(* IEC 61131-3 sources: daoli-st-library/DL_Motion (part 10) *)

(* ---- FB_DL_AxisTorqueRippleWatch.st ---- *)
(*
  Name        : FB_DL_AxisTorqueRippleWatch
  Category    : DL_Motion
  Version     : 1.0.0
  Purpose     : 轴转矩纹波监视：匀速段窗内峰峰值/均值占比与峰间隔规律性双判据，识别机械卡滞与联轴器异常；/ Axis torque ripple watch: peak-to-mean ripple ratio and peak-interval regularity in a steady-speed window to identify mechanical sticking and coupling anomalies
  溯源        : 借 plcopen-motion 的运动诊断组织，clean-room 实现
  Boundary    : ① 只在匀速段采样（|速度 - 速度命令| < 容差 且 速度 > 最低速），运动相位闸（容差/最低速域 > 0）；
                ② 波动幅度 = 窗内峰峰值 / 均值占比判据，均值近零时占比出口置 0 + bInvalid（除零前置）；
                ③ 周期性判据 = 峰间隔极差 < 阈（机械卡滞特征），需窗内 >= 3 个局部峰才判；
                ④ 非有限扭矩该拍不入窗（窗保持不滑动，防污染统计）；
                ⑤ 本件为诊断观测层，不干预轴指令输出（属主边界，零控制量引脚）；
                ⑥ 窗长 32 固定常量，窗内统计每趟全量重算防陈旧（R227）。
*)
TYPE E_DL_TrwState :
(
    eIdle  := 0,                             (* 未使能（窗清空） / Disabled, window cleared *)
    eRun   := 10,                            (* 纹波监视运行 / Watching *)
    eFault := 90                             (* 故障锁存相 / Fault latched *)
);
END_TYPE

TYPE E_DL_TrwCause :
(
    eNone      := 0,                         (* 无成因 / No cause *)
    eCfgIllegal:= 1,                        (* 组态非法：容差/最低速/阈值/周期越域 / Illegal config *)
    ePhaseBad  := 2                         (* 非法相位兜底 / Illegal phase fallback *)
);
END_TYPE

FUNCTION_BLOCK FB_DL_AxisTorqueRippleWatch
VAR_INPUT
    fTorque  : REAL := 0.0;                  (* 轴转矩反馈 [Nm] / Axis torque feedback *)
    fVel     : REAL := 0.0;                 (* 轴实际速度 [mm/s] / Actual velocity *)
    fVelCmd  : REAL := 0.0;                 (* 轴速度命令（匀速判据基准）[mm/s] / Velocity command *)
    fVelTol  : REAL := 5.0;                  (* 匀速判据容差，域 > 0 [mm/s] / Steady-speed tolerance *)
    fVelMin  : REAL := 10.0;                 (* 最低采样速度，域 > 0 [mm/s] / Minimum sampling speed *)
    fTqLimRip: REAL := 10.0;                 (* 纹波占比报警阈，域 > 0 [%] / Ripple ratio limit *)
    fGapSpreadMax: REAL := 0.05;             (* 峰间隔极差阈，域 > 0 [s] / Gap spread limit *)
    tSample  : TIME := T#10MS;               (* 采样周期，域 > T#0S [ms] / Sampling period *)
    bEnable  : BOOL := TRUE;                 (* 使能 [-] / Enable *)
    bReset   : BOOL := FALSE;                (* 复位命令，上升沿清窗与故障 [-] / Reset command *)
END_VAR
VAR_OUTPUT
    fRipplePct: REAL;                        (* 纹波占比出口 = 峰峰值 / |均值| × 100 [%] / Ripple ratio outlet *)
    bRippleHigh: BOOL;                       (* 纹波超阈判据出口 [-] / Ripple high verdict *)
    bPeriodic: BOOL;                         (* 周期性卡滞特征出口（>= 3 峰且间隔规律）[-] / Periodic sticking verdict *)
    bInvalid : BOOL;                         (* 本拍统计无效指示（均值近零/样本不足）[-] / Invalid indicator *)
    eState   : E_DL_TrwState;                (* 状态出口 / State outlet *)
    eCause   : E_DL_TrwCause;                (* 故障成因出口（R190 归因唯一） / Fault cause outlet *)
    bError   : BOOL;                         (* 故障锁存标志 [-] / Fault latch flag *)
END_VAR
VAR
    _eState : E_DL_TrwState := E_DL_TrwState.eIdle;  (* 内部相位（CASE 唯一写入目标） / Internal phase *)
    _eCause : E_DL_TrwCause := E_DL_TrwCause.eNone;  (* 成因锁存量 / Latched cause *)
    rtReset : R_TRIG;                        (* 复位沿实例，段 0 无条件调用 / Reset edge instance *)
    _bFault : BOOL;                          (* 故障锁存位 / Latched fault bit *)
    _bCfgBad: BOOL;                          (* 组态非法当拍量 / Illegal config this scan *)
    _bFin   : BOOL;                          (* 扭矩有限性当拍量（边界④） / Torque finiteness *)
    _bSteady: BOOL;                          (* 匀速段当拍判据（边界①） / Steady-speed verdict *)
    _aWin   : ARRAY[1..32] OF REAL;          (* 扭矩滑窗（线性平移式）[Nm] / Torque sliding window *)
    _nFill  : INT;                           (* 窗填充数 [点] / Window fill count *)
    _i      : INT;                           (* 窗扫描游标 [点] / Window scan cursor *)
    _fMean  : REAL;                          (* 窗均值中间量 [Nm] / Window mean *)
    _fPk    : REAL;                          (* 窗峰值中间量 [Nm] / Window peak *)
    _fTr    : REAL;                          (* 窗谷值中间量 [Nm] / Window trough *)
    _fSum   : REAL;                          (* 窗求和中间量 [Nm] / Window sum *)
    _nPkN   : INT;                           (* 本趟局部峰计数 [个] / Local peak count *)
    _nLastPk: INT;                           (* 上一峰样本序号（间隔派生）[点] / Last peak index *)
    _aGap   : ARRAY[1..4] OF REAL;           (* 最近峰间隔表（秒值）[s] / Recent peak gaps *)
    _nGapN  : INT;                           (* 已存间隔数 [个] / Stored gap count *)
    _fGapMax: REAL;                          (* 间隔极差上界中间量 [s] / Gap spread upper *)
    _fGapMin: REAL;                          (* 间隔极差下界中间量 [s] / Gap spread lower *)
    _fDtSec : REAL;                          (* 采样周期秒值，域 > eps [s] / Sampling period seconds *)
    _bPerI  : BOOL;                          (* 周期性判据内部量 / Periodic verdict internal *)
END_VAR
VAR CONSTANT
    DL_TRW_NMAX : INT   := 32;               (* 滑窗容量（固定常量，边界⑥）[点] / Window capacity *)
    DL_TRW_NMIN : INT   := 8;                (* 统计生效最少样本数（防小样本误判）[点] / Minimum samples *)
    DL_TRW_NPKMIN: INT  := 3;                (* 周期性判据最少峰数（边界③）[个] / Minimum peaks *)
    DL_TRW_EPS  : REAL  := 1.0E-6;           (* 判零容差 [-] / Epsilon *)
END_VAR

(* —— 段 0：当拍判据派生 + 实例无条件刷新（R228A） —— *)
_fDtSec := TIME_TO_LREAL(tSample) / 1000.0;              (* 采样周期秒化（除子常量 1000） / Sampling period seconds *)
_bCfgBad := (fVelTol <= DL_TRW_EPS) OR (fVelMin <= DL_TRW_EPS)           (* 匀速容差/最低速正域闸（边界①） / Tolerance and speed gates *)
            OR (fTqLimRip <= DL_TRW_EPS) OR (fGapSpreadMax <= DL_TRW_EPS)   (* 报警阈正域闸（边界②③） / Verdict limit gates *)
            OR NOT (tSample > T#0S);                     (* 采样周期正域闸 / Sampling gate *)
rtReset(CLK := bReset);                                  (* 复位沿每拍必调 / Reset edge every scan *)
_bFin := (fTorque = fTorque) AND ((fTorque - fTorque) = (fTorque - fTorque));   (* 扭矩 NaN 自反 + Inf 差判闸（边界④） / Torque NaN and Inf gate *)
_bSteady := (ABS(fVel - fVelCmd) < fVelTol) AND (fVel > fVelMin);        (* 匀速段判据：速度差容差内且高于最低速（边界①） / Steady-speed verdict *)

(* —— 段 1：单拍量预清零（R107；出口在段 4 每趟重算前预置确定值） —— *)
fRipplePct := 0.0;                                       (* 占比出口预清（无效拍默认 0） / Ripple preset zero *)
bRippleHigh := FALSE;                                    (* 超阈出口预清 / High preset *)
bPeriodic := FALSE;                                      (* 周期性出口预清 / Periodic preset *)
bInvalid := FALSE;                                       (* 无效指示预清 / Invalid preset *)
_bPerI := FALSE;                                         (* 周期性内部量预清（R227） / Periodic internal clear *)
_nPkN := 0;                                              (* 峰计数每趟重置 / Peak count reset *)
_nLastPk := 0;                                           (* 峰序号快照重置 / Peak index reset *)
_nGapN := 0;                                             (* 间隔表计数每趟重算 / Gap count reset *)
_fGapMax := 0.0;                                         (* 极差上界重置 / Spread upper reset *)
_fGapMin := 0.0;                                         (* 极差下界重置 / Spread lower reset *)

(* —— 段 2：复位沿处理（作用域：清故障 + 清窗 + 迁 eIdle，R283 逐项声明） —— *)
IF rtReset.Q THEN
    _bFault := FALSE;                                    (* 清故障锁存 / Clear fault *)
    _eCause := E_DL_TrwCause.eNone;                      (* 清成因 / Clear cause *)
    FOR _i := 1 TO DL_TRW_NMAX DO
        _aWin[_i] := 0.0;                                (* 清滑窗 / Clear window *)
    END_FOR
    FOR _i := 1 TO 4 DO
        _aGap[_i] := 0.0;                                (* 清间隔表 / Clear gap table *)
    END_FOR
    _nFill := 0;                                         (* 清窗填充数 / Clear fill *)
    fRipplePct := 0.0;                                   (* 清占比出口 / Clear ripple outlet *)
    _eState := E_DL_TrwState.eIdle;                      (* 迁未使能相 / Back to idle *)
END_IF

(* —— 段 3：组态故障锁存（锁存至复位沿，R189） —— *)
IF _bCfgBad AND NOT _bFault THEN
    _bFault := TRUE;                                     (* 锁存故障位 / Latch fault *)
    _eCause := E_DL_TrwCause.eCfgIllegal;                (* 成因：组态非法 / Cause illegal config *)
    _eState := E_DL_TrwState.eFault;                     (* 同步迁故障相 / Migrate to fault *)
END_IF

(* —— 段 4：CASE 主状态机（ELSE 兜底迁 eFault，红线 6） —— *)
CASE _eState OF
    E_DL_TrwState.eIdle:                                 (* 未使能：窗清空出口确定值 / Idle *)
        FOR _i := 1 TO DL_TRW_NMAX DO
            _aWin[_i] := 0.0;                            (* 失能清滑窗 / Disabled clear window *)
        END_FOR
        _nFill := 0;                                     (* 失能清填充数 / Disabled clear fill *)
        IF bEnable AND NOT _bFault THEN
            _eState := E_DL_TrwState.eRun;               (* 进入监视相 / Enter watching *)
        END_IF
    E_DL_TrwState.eRun:                                  (* 监视相：匀速闸采样 + 全窗重算 / Watching *)
        IF NOT bEnable THEN
            _eState := E_DL_TrwState.eIdle;              (* 失能回未使能 / Back to idle *)
        ELSE
            IF _bSteady AND _bFin AND (_fDtSec > DL_TRW_EPS) THEN   (* 匀速闸 + 有限闸 + 周期闸（边界①④） / Sampling gates *)
                IF _nFill < DL_TRW_NMAX THEN
                    _nFill := _nFill + 1;                (* 填充数递进（写入点域内） / Fill advance *)
                    _aWin[_nFill] := fTorque;            (* 样本入窗 / Sample into window *)
                ELSE
                    FOR _i := 1 TO DL_TRW_NMAX - 1 DO
                        _aWin[_i] := _aWin[_i + 1];      (* 满窗线性平移（有界循环） / Shift window *)
                    END_FOR
                    _aWin[DL_TRW_NMAX] := fTorque;       (* 新样本入窗尾 / Sample into tail *)
                END_IF
            END_IF                                       (* 不满足闸：本拍不入窗（窗保持，边界①④） *)
            IF _nFill >= DL_TRW_NMIN THEN                (* 统计生效下限（防小样本误判） / Statistics gate *)
                _fSum := 0.0; _fPk := _aWin[1]; _fTr := _aWin[1];   (* 均值/峰谷初值（R227） / Init mean peak trough *)
                FOR _i := 1 TO _nFill DO
                    _fSum := _fSum + _aWin[_i];          (* 窗求和 / Window sum *)
                    IF _aWin[_i] > _fPk THEN
                        _fPk := _aWin[_i];               (* 窗峰值刷新 / Peak update *)
                    END_IF
                    IF _aWin[_i] < _fTr THEN
                        _fTr := _aWin[_i];               (* 窗谷值刷新 / Trough update *)
                    END_IF
                END_FOR
                _fMean := _fSum / INT_TO_REAL(_nFill);   (* 窗均值（除子 = 填充数 >= 8） / Window mean *)
                IF ABS(_fMean) > DL_TRW_EPS THEN
                    fRipplePct := (_fPk - _fTr) / ABS(_fMean) * 100.0;   (* 纹波占比（除子已过闸，边界②） / Ripple ratio *)
                    bRippleHigh := fRipplePct > fTqLimRip;   (* 占比超阈判据（直比阈值） / Ripple high verdict *)
                ELSE
                    fRipplePct := 0.0;                   (* 均值近零：占比出口 0（除零前置，边界②） / Zero ratio *)
                    bInvalid := TRUE;                    (* 无效指示 / Invalid indicator *)
                END_IF
                FOR _i := 2 TO _nFill - 1 DO             (* 局部峰检测（内点扫描，边界③） / Local peak scan *)
                    IF (_aWin[_i] > _aWin[_i - 1]) AND (_aWin[_i] > _aWin[_i + 1]) AND (_aWin[_i] > _fMean) THEN
                        _nPkN := _nPkN + 1;              (* 局部峰计数 / Peak count *)
                        IF _nLastPk >= 1 THEN
                            _nGapN := _nGapN + 1;        (* 间隔数净额 +1 / Gap count *)
                            IF _nGapN > 4 THEN
                                _aGap[1] := _aGap[2]; _aGap[2] := _aGap[3]; _aGap[3] := _aGap[4];   (* 间隔表平移 / Shift gaps *)
                                _nGapN := 4;             (* 间隔表封顶 / Gap cap *)
                            END_IF
                            _aGap[_nGapN] := INT_TO_REAL(_i - _nLastPk) * _fDtSec;   (* 间隔秒值入表 / Gap into table *)
                        END_IF
                        _nLastPk := _i;                  (* 峰序号快照 / Peak index snapshot *)
                    END_IF
                END_FOR
                IF _nGapN >= 2 THEN                      (* >= 3 峰（2 个间隔）才判（边界③） / Peak count gate *)
                    _fGapMax := _aGap[1]; _fGapMin := _aGap[1];   (* 极差初值 / Spread init *)
                    FOR _i := 2 TO _nGapN DO
                        IF _aGap[_i] > _fGapMax THEN
                            _fGapMax := _aGap[_i];       (* 间隔上界刷新 / Gap upper *)
                        END_IF
                        IF _aGap[_i] < _fGapMin THEN
                            _fGapMin := _aGap[_i];       (* 间隔下界刷新 / Gap lower *)
                        END_IF
                    END_FOR
                    _bPerI := (_fGapMax - _fGapMin) < fGapSpreadMax;   (* 间隔规律性判据（边界③） / Regularity verdict *)
                END_IF
                bPeriodic := _bPerI;                     (* 周期性出口 / Periodic outlet *)
            ELSE
                bInvalid := TRUE;                        (* 样本不足：统计无效（确定值） / Not enough samples *)
            END_IF
        END_IF
    E_DL_TrwState.eFault:                                (* 故障相：冻结保持，仅复位沿出 / Fault *)
        ;                                                (* 锁存回放（R28） / Replay from latch *)
    ELSE                                                 (* 非法相位兜底迁安全态 / Illegal phase fallback *)
        _eState := E_DL_TrwState.eFault; _bFault := TRUE;    (* 迁故障相 + 同步锁存 / To fault and latch *)
        _eCause := E_DL_TrwCause.ePhaseBad;              (* 成因：非法相位 / Cause illegal phase *)
END_CASE

(* —— 段 5：出口映射（bError/eState 同源，R191） —— *)
bError := _bFault;                                       (* 故障标志镜像 / Fault flag mirror *)
eState := _eState;                                       (* 状态出口 / State outlet *)
eCause := _eCause;                                       (* 成因出口 / Cause outlet *)
END_FUNCTION_BLOCK

(* ---- FB_DL_AxisTorqueWatch.st ---- *)
(*
  组件名 Component   : FB_DL_AxisTorqueWatch
  子库 Sublibrary    : DL_Motion
  版本 Version       : 1.0.0
  兼容性 Platform    : CODESYS 3.5 / TwinCAT 3 / 汇川 InoProShop / Machine Expert（仅 Standard.library）
  功能 Function      : 轴转矩趋势监视（与 FB_DL_TorqueLimitControl 分工：控 vs 监）：
                       1) 带域判据：转矩超上带限持续 tConfirmWin → 预警（bWarn）；
                       2) 趋势斜率判据：周期窗（tSlopeWin 自复触）两端采样，斜率
                       fSlopeNmS = (本端 - 上端) / 窗长，斜率超限 → 预警；
                       3) 堵转分级：转矩超上带限 且 轴速近零 持续 tStallTo → bStall；
                       4) 三判据各带独立确认窗，互不共用计时实例（R190 归因唯一）。
  边界 Boundary      : ① 监视件只出分级诊断位，不接管转矩控制输出；
                       ② 周期窗计时用 IN := bEnable AND NOT tonSlopeWin.Q 自复触
                       （R188 错峰周期窗范式，禁外部沿清零）；
                       ③ 斜率除法前置域闸：tSlopeWin <= T#0S 判组态非法；
                       ④ 非有限值（NaN 自反 + 无穷差值自减）判输入非法锁存；
                       ⑤ 故障锁存解除唯一路径 = bReset 上升沿（输入引脚，恒可达）；
                       ⑥ 无全局变量引用、无外部变量声明、无物理地址寻址。
  依赖 Depends       : Standard.library（R_TRIG / TON）
  溯源 Origin        : 道莅自研 clean-room（参考 t2-4-s7-motion 监视分类与参数域，
                       零代码行复制）
  码位 Code          : 16#04_0_A9
  码表 Error codes（Motion 格 04_0_A9，单轨：故障 0x02A9 / 信息 0x01A9 / 0x03A9）:
    16#0004_02A9 故障级：组态非法或输入非有限，锁存至 bReset 上升沿
    16#0004_01A9 信息级：预警进入沿（bWarn 由 FALSE 转 TRUE 拍）
    16#0004_05A9 信息级：堵转检出沿（bStall 由 FALSE 转 TRUE 拍；子道 05 为 03 道撞车顺延勘误）
  修订历史 Revision  :
    2026-11-19  v1.0.0  R44 首版（批次 2 · 序号 6）
*)

TYPE E_DL_AtwState :
(
    eIdle  := 0,    // 空闲：未使能 / Idle, not enabled
    eRun   := 10,   // 监视运行：三判据并行 / Running, three criteria active
    eFault := 90    // 故障：组态/输入锁存 / Fault, latched
);
END_TYPE

FUNCTION_BLOCK FB_DL_AxisTorqueWatch
VAR_INPUT
    bEnable    : BOOL;                     // 使能（电平）[-] / Enable
    bReset     : BOOL;                     // 上升沿清故障锁存 [-] / Reset edge
    fTorqueNm  : REAL;                     // 实测转矩 [牛·米] / Measured torque
    fVelMmS    : REAL;                     // 轴实际速度 [mm/s] / Axis velocity
    fBandHiNm  : REAL := 10.0;             // 转矩上带限 [牛·米] / Torque band ceiling
    fBandLoNm  : REAL := 1.0;              // 转矩下带限 [牛·米] / Torque band floor
    fSlopeLimNmS: REAL := 5.0;             // 趋势斜率限值 [牛·米/秒] / Trend slope limit
    fVelNearZeroMmS: REAL := 0.5;          // 堵转判近零速度阈 [mm/s] / Near-zero velocity threshold
    tConfirmWin: TIME := T#2S;             // 带域预警确认窗 [毫秒] / Band confirm window
    tSlopeWin  : TIME := T#1S;             // 趋势斜率测量窗 [毫秒] / Slope measurement window
    tStallTo   : TIME := T#3S;             // 堵转确认窗 [毫秒] / Stall confirm window
END_VAR
VAR_OUTPUT
    bInBand    : BOOL;                     // 转矩在带内电平 [-] / Torque in-band level
    bWarn      : BOOL;                     // 预警电平（带域或斜率越限确认后）[-] / Warning level
    bStall     : BOOL;                     // 堵转电平 [-] / Stall level
    fSlopeNmS  : REAL;                     // 实测趋势斜率 [牛·米/秒] / Measured slope
    eState     : E_DL_AtwState;            // 状态出口，段尾单点映射 / State outlet
    bError     : BOOL;                     // 故障锁存标志 [-] / Fault latch flag
    uErrId     : UDINT;                    // 事件码，0 = 无事件 / Event code
END_VAR
VAR
    rtReset    : R_TRIG;                   // 复位沿实例，段 0 无条件刷新 / Reset edge
    rtWarn     : R_TRIG;                   // 预警进入沿实例，段 0 无条件刷新 / Warn entry edge
    rtStall    : R_TRIG;                   // 堵转进入沿实例，段 0 无条件刷新 / Stall entry edge
    tonBandWin : TON;                      // 带域确认窗（专用确认窗命名） / Band confirm timer
    tonStallTo : TON;                      // 堵转确认窗（专用超时件命名（R228A 豁免）） / Stall timer
    tonSlopeWin: TON;                      // 斜率周期窗（自复触，R188） / Slope window timer
    _eState    : E_DL_AtwState := E_DL_AtwState.eIdle;   // 内部相位（CASE 唯一写入目标）/ Internal phase
    _bBandHi   : BOOL;                     // 带域越限当拍量 [-] / Band breach flag
    _bStallCond: BOOL;                     // 堵转条件当拍量 [-] / Stall condition flag
    _fTorqueSnap: REAL;                    // 窗始转矩快照 [牛·米] / Window-start torque snapshot
    _bSnapPend : BOOL;                     // 快照待取标志 [-] / Snapshot pending flag
    _bFault    : BOOL;                     // 故障锁存位（锁存量） / Latched fault bit
    _uFault    : UDINT;                    // 故障码锁存（锁存量） / Latched fault code
    _bCfgBad   : BOOL;                     // 组态非法当拍量 [-] / Config illegal flag
    _bNonFin   : BOOL;                     // 输入非有限当拍量 [-] / Non-finite input flag
END_VAR
VAR CONSTANT
    DL_SLOPE_EPS: REAL := 1.0E-9;          // 斜率判零容差 [牛·米/秒] / Slope tolerance
    DL_WIN_EPS  : REAL := 1.0E-3;          // 窗长秒值下限 [秒] / Window seconds floor
    DL_ABS_MAX  : REAL := 1.0E30;          // 有限值判定上界 [工程单位] / Finite bound
    DL_ZERO     : REAL := 0.0;             // 零常量 [工程单位] / Zero constant
    DL_MS_PER_S : REAL := 1000.0;          // 毫秒 → 秒换算系数 [毫秒/秒] / Milliseconds per second
END_VAR

(* —— 段 0｜沿与定时器每拍无条件刷新（禁置于 IF/CASE 内） —— *)
_bBandHi    := (fTorqueNm > fBandHiNm) OR (fTorqueNm < fBandLoNm);   // 带域越限当拍判据
_bStallCond := (fTorqueNm > fBandHiNm) AND (ABS(fVelMmS) < fVelNearZeroMmS);
rtReset    (CLK := bReset);
rtWarn     (CLK := bWarn);
rtStall    (CLK := bStall);
tonBandWin (IN := (_eState = E_DL_AtwState.eRun) AND _bBandHi AND (NOT _bFault), PT := tConfirmWin);
tonStallTo (IN := (_eState = E_DL_AtwState.eRun) AND _bStallCond AND (NOT _bFault), PT := tStallTo);
tonSlopeWin(IN := (_eState = E_DL_AtwState.eRun) AND (NOT _bFault) AND (NOT tonSlopeWin.Q),
            PT := tSlopeWin);            // 自复触周期窗：Q 拍断开一拍，下拍重启（R188）

(* —— 段 1｜瞬时量预清零（锁存量 _bFault/_uFault/bWarn/bStall/_fTorqueSnap 不入清单） —— *)
uErrId   := 16#0000_0000;
_bCfgBad := FALSE;
_bNonFin := FALSE;

(* —— 段 2｜复位沿：故障一次性清干净，相位回空闲，诊断位复归 —— *)
IF rtReset.Q THEN
    _bFault  := FALSE;
    _uFault  := 16#0000_0000;
    bWarn    := FALSE;
    bStall   := FALSE;
    fSlopeNmS:= DL_ZERO;
    _eState  := E_DL_AtwState.eIdle;
END_IF

(* —— 段 3｜组态闸与非有限判据 —— *)
IF (fBandHiNm <= fBandLoNm) OR (tConfirmWin = T#0S) OR (tSlopeWin = T#0S)
   OR (tStallTo = T#0S) OR (fVelNearZeroMmS <= DL_ZERO) THEN
    _bCfgBad := TRUE;
END_IF
IF (fTorqueNm <> fTorqueNm) OR ((fTorqueNm - fTorqueNm) <> DL_ZERO)
   OR (fVelMmS <> fVelMmS) OR ((fVelMmS - fVelMmS) <> DL_ZERO) THEN
    _bNonFin := TRUE;
END_IF

(* —— 段 4｜主状态机：三态全覆盖 + ELSE 兜底 —— *)
CASE _eState OF

E_DL_AtwState.eIdle:
    bInBand := FALSE;
    IF bEnable AND (NOT _bCfgBad) AND (NOT _bNonFin) THEN
        _fTorqueSnap := fTorqueNm;       // 窗始快照初始化
        _bSnapPend   := FALSE;
        _eState := E_DL_AtwState.eRun;
    ELSIF bEnable AND (_bCfgBad OR _bNonFin) THEN
        _bFault := TRUE;
        _uFault := 16#0004_02A9;
        bError  := TRUE;
        _eState := E_DL_AtwState.eFault;
    END_IF

E_DL_AtwState.eRun:
    IF NOT bEnable THEN
        bInBand := FALSE;
        bWarn   := FALSE;
        bStall  := FALSE;
        _eState := E_DL_AtwState.eIdle;  // 使能撤销回空闲
    ELSE
        bInBand := NOT _bBandHi;
        (* 斜率测量：Q 拍收口，快照按窗复归（除数 = 窗长秒值，组态闸已保证 > 0） *)
        IF tonSlopeWin.Q THEN
            IF NOT _bSnapPend THEN
                fSlopeNmS := (fTorqueNm - _fTorqueSnap)
                             / MAX(TIME_TO_REAL(tSlopeWin) / DL_MS_PER_S, DL_WIN_EPS);
                IF ABS(fSlopeNmS) < DL_SLOPE_EPS THEN
                    fSlopeNmS := DL_ZERO;    // 斜率近零归零
                END_IF
                _bSnapPend := TRUE;
            END_IF
            _fTorqueSnap := fTorqueNm;
            _bSnapPend   := FALSE;
        END_IF
        (* 分级判据：带域或斜率任一确认 → 预警；带域 + 近零速度确认 → 堵转 *)
        IF _bNonFin THEN
            _bFault := TRUE;             // 输入非有限：运行中锁存
            _uFault := 16#0004_02A9;
            bError  := TRUE;
            bWarn   := FALSE;
            bStall  := FALSE;
            _eState := E_DL_AtwState.eFault;
        ELSE
            bWarn := (NOT _bFault) AND (tonBandWin.Q OR (ABS(fSlopeNmS) > fSlopeLimNmS));
            bStall := (NOT _bFault) AND tonStallTo.Q;
            IF rtWarn.Q THEN
                uErrId := 16#0004_01A9;  // 信息级：预警进入沿
            END_IF
            IF rtStall.Q THEN
                uErrId := 16#0004_05A9;  // 信息级：堵转检出沿（子道 05 勘误顺延）
            END_IF
        END_IF
    END_IF

E_DL_AtwState.eFault:
    bError := TRUE;                      // 故障相驻留：诊断位冻结，只认复位沿（段 2 迁出）
    ;                                    // （冻结语义：bWarn/bStall 保持复位沿前值由段 2 归零）

ELSE
    _bFault := TRUE;                     // 兜底：非法相位锁存
    _uFault := 16#0004_02A9;
    bError  := TRUE;
    _eState := E_DL_AtwState.eFault;
END_CASE

(* —— 段 5｜状态出口单点映射 —— *)
eState := _eState;
END_FUNCTION_BLOCK

(* ---- FB_DL_AxisVelocityMove.st ---- *)
(*==============================================================================
 * 组件名称 (Component)  : FB_DL_AxisVelocityMove
 * 所属子库 (Sublibrary) : DL_Motion
 * 当前版本 (Version)    : 1.0.0
 * 组件分类 (Category)   : 功能块（FUNCTION_BLOCK）· 单轴速度模式与动态变速封装 · 工艺上层件
 * 兼容性   (Platform)   : CODESYS 3.5 / TwinCAT 3 / 汇川 InoProShop / Schneider
 *                         Machine Expert；仅依赖 Standard.library（R_TRIG /
 *                         F_TRIG / MIN / MAX / ABS），零厂商方言
 * 接口依赖 (Depends)    : I_DL_MotionAxis / E_DL_AxisState（既有契约，Round 05）
 * 功能描述 (Function)   : 单轴速度模式（MC_MoveVelocity 语义）与动态变速控制
 *                         封装。经轴接口引用驱动轴体：指令电平生效，TRUE=运行
 *                         / FALSE=受控停止；运行中变更 fVelocity 即为改速请求
 *                         （轴接口连续运动改速语义，改速而非重启），bDynamicRetarget
 *                         使能时自动重发；速度上限独立钳位，越限置信息级。
 * 设计要点 (Key notes)  : ① 指令上升沿门禁：轴待机态受理运行、连续运动态受理
 *                           改速；其余态请求不被受理 → 信息级 0004_0107；
 *                         ② 动态改速：连续运动中 |fVelocity − 上次已发值| 超
 *                           容差即重发 MoveVelocity（改速语义），指令被拒 →
 *                           0004_0230 故障级锁存；
 *                         ③ 下降沿 → 轴受控停止（MC_Stop 语义）；
 *                         ④ 参数门禁（fAcc 非正值/非有限值）→ 信息级 0004_0106
 *                           （与 FB_DL_AxisHomingSeq/FB_DL_AxisRelativeMove
 *                           同码同义：参数门禁拒绝，共用留档）；
 *                         ⑤ 本块为事件型 + 轮询状态组件，免首扫（R23）。
 * 开源溯源 (Origin)     : 原创实现（参考 PLCopen Part 1-6 MC_MoveVelocity 公开
 *                         语义与西门子 Motion Control 对象语义，clean-room）。
 *                         仅提取公开指令动词、参数域与改速语义；实现与命名
 *                         100% 自有，未参考任何厂商源码行。
 * 验收向量 (Acceptance) :
 *   V1 启动-停止链：bCmdStart 上升沿→轴进连续运动；下降沿→受控停止；
 *   V2 运行中改速：fVelocity 50→-30（含反向）→ 自动重发改速，轴不重启；
 *   V3 改速被拒：轴受控停止中发改速请求 → 信息级 0004_0107，轴不受扰；
 *   V4 速度钳位：|fVelocity|=5000 > fVelMax=1000 → 钳位至 1000 + 信息级；
 *   V5 轴故障中断：运行中轴故障反馈 → 0004_0230 锁存，bBusy 退出。
 * 故障码表 (Error codes):
 *   16#0004_0106【信息级】参数门禁拒绝（三块同码同义，共用留档）；
 *   16#0004_0107【信息级】改速请求不被受理/速度钳位提示（规格外补充子义，
 *   R11 留档）；16#0004_0230【故障级】指令被拒/轴故障中断（锁存）；
 *   16#0004_0201【故障级】非法状态兜底（沿用族码，与 FB_DL_SingleAxis 同码
 *   同义，复用留档）。
 * 修订历史 (Revision)   :
 *   2026-11-15  v1.0.0  首版入库（Round 06 · DL_Motion 回零/运动族）
 *============================================================================*)

(*-----------------------------------------------------------------------------
 * 调用示例 (Instance guide)：
 *   fbVel.iAxis := fbAxis;                        // 接口依赖注入
 *   fbVel(bCmdStart := bRunSwitch, fVelocity := fSetVel, // 周期调用
 *         fAcc := 2000.0, bDynamicRetarget := TRUE, fVelMax := 1000.0);
 *   电平语义：bRunSwitch 断开即受控减速停车，无需上层编排停止时序；
 *   改速只需改 fVelocity 输入值，块自动差值比较后重发改速指令。
 *----------------------------------------------------------------------------*)

(*-----------------------------------------------------------------------------
 * 常见误用与现场提示 (Field notes)：
 *   1 bCmdStart 电平语义：FALSE 即停车并退出速度模式，不要用脉冲；
 *     需要脉冲语义的工位在上层自锁存。
 *   2 改速容差为固定值（0.001 mm/s），HMI 微调速度时每次变化都会重发；
 *     高频改速场景请在上层做死区滤波，避免指令流量放大。
 *   3 轴限位停车后 bCmdStart 仍为 TRUE 时本块会自动重新发起（电平需求
 *     语义）；不希望自动重启的工位在限位联动层断开 bCmdStart。
 *----------------------------------------------------------------------------*)

(*-----------------------------------------------------------------------------
 * 枚举: E_DL_VelStep（归属 DL_Motion，与 FB_DL_AxisVelocityMove 同文件）
 * 含义: 速度模式内部步进枚举（本块私有配套，外部仅作诊断参考）。
 *----------------------------------------------------------------------------*)
{attribute 'strict'}
{attribute 'qualified_only'}
TYPE E_DL_VelStep :
(
    eIdle    := 0,    // 空闲：等待启动沿 / Idle: waiting for start edge
    eRunning := 10    // 运行：轮询轴状态并处理动态改速 / Running: polling axis and retargeting
) UINT;
END_TYPE

FUNCTION_BLOCK FB_DL_AxisVelocityMove
VAR_INPUT
    bCmdStart        : BOOL := FALSE;   // 速度运行指令（Velocity start command），电平生效：TRUE=运行 / FALSE=受控停止
    fVelocity        : REAL := 0.0;     // 目标速度（Target velocity）[mm/s]，带符号，负值=负向；运行中变更即为改速请求
    fAcc             : REAL := 1000.0;  // 加减速度（Acceleration）[mm/s²]，正值，默认 1000.0
    bDynamicRetarget : BOOL := FALSE;   // 动态改速使能（Dynamic retarget），TRUE=连续运动中速度变化自动改速
    fVelMax          : REAL := 1000.0;  // 速度上限（Velocity limit）[mm/s]，|fVelocity| 超限钳位并置信息级
END_VAR
VAR_IN_OUT
    iAxis            : I_DL_MotionAxis; // 轴接口引用（Axis reference），由上层注入实现块实例
END_VAR
VAR_OUTPUT
    bBusy            : BOOL := FALSE;   // 速度模式激活（Velocity mode active）
    bActive          : BOOL := FALSE;   // 轴处于连续运动态（Axis in continuous motion），轮询派生
    uErrorId         : UDINT := 0;      // 末次事件码（Last error code），段位 16#0004_xxxx
END_VAR
VAR
    eStep            : E_DL_VelStep := E_DL_VelStep.eIdle; // 内部步进状态（Internal step state）
    bFaultLatch      : BOOL := FALSE;   // 故障锁存标志（Fault latch），0004_0230 锁存载体
    bParamOk         : BOOL := FALSE;   // 参数门禁通过标志（Parameter gate pass flag），逐拍重算
    fVelEff          : REAL := 0.0;     // 本拍钳位后的目标速度（Clamped target velocity）[mm/s]
    fVelSent         : REAL := 0.0;     // 上次已发轴指令速度（Last issued velocity）[mm/s]，改速差值比较基准
    fVelLim          : REAL := 1000.0;  // 生效速度上限（Effective velocity limit）[mm/s]，非有限值兜底
    fAccEff          : REAL := 1000.0;  // 生效加减速度（Effective acceleration）[mm/s²]，防除零兜底
    rtrigStart       : R_TRIG;          // 启动指令上升沿（Rising edge of start command）
    ftrigStart       : F_TRIG;          // 启动指令下降沿（Falling edge of start command）
END_VAR
VAR CONSTANT
    DL_VEL_INF_MAX   : REAL := 1.0E30;  // 有限值判定幅值上限（Finite-value magnitude bound）[mm/s 或 mm/s²]
    DL_VEL_EPS       : REAL := 1.0E-6;  // 浮点判零容差（Float zero tolerance）
    DL_VEL_TGT_TOL   : REAL := 1.0E-3;  // 改速差值容差（Retarget delta tolerance）[mm/s]，超过才重发改速
    DL_VEL_PAR_FLOOR : REAL := 1.0E-3;  // 加速度参数下限（Acceleration floor）[mm/s²]
END_VAR

// 段 1｜沿检测无条件周期刷新（R7 红线，严禁置于分支内）
rtrigStart(CLK := bCmdStart);
ftrigStart(CLK := bCmdStart);

// 段 2｜接口引用有效性防御：未注入轴引用则清输出退出（不产生误动作）
IF iAxis = 0 THEN
    bBusy := FALSE;
    bActive := FALSE;
    RETURN;
END_IF

// 段 3｜参数门禁逐拍重算（公约 0.8）：非法仅封锁启动（信息级 0004_0106），运行中不中断
bParamOk := (fAcc = fAcc) AND (fAcc <= DL_VEL_INF_MAX) AND (fAcc > DL_VEL_PAR_FLOOR);
IF (fVelMax = fVelMax) AND (fVelMax > DL_VEL_PAR_FLOOR) AND (fVelMax <= DL_VEL_INF_MAX) THEN
    fVelLim := fVelMax;                          // 合法速度上限直通 [mm/s]
ELSE
    fVelLim := 1000.0;                           // 非法上限兜底 [mm/s]
    uErrorId := 16#0004_0106;                    // 信息级：参数兜底修复提示
END_IF
fAccEff := MAX(fAcc, DL_VEL_PAR_FLOOR);          // 生效加速度下限兜底 [mm/s²]，防除零

// 段 4｜事件码管理（R15）：瞬时码逐拍重算，锁存码仅在新启动沿解除
IF NOT bFaultLatch THEN
    uErrorId := 0;
END_IF

// 段 5｜下降沿受控停车（电平语义：FALSE=停止；全局处理，任何态均生效）
IF ftrigStart.Q THEN
    iAxis.Stop();                                // 受控减速停车（MC_Stop 语义）
    bBusy := FALSE;
    IF eStep = E_DL_VelStep.eRunning THEN
        eStep := E_DL_VelStep.eIdle;             // 退出速度模式，等待下次启动沿
    END_IF
END_IF

// 段 6｜运行中轴故障中断（优先于状态机，锁存 R15）
IF (eStep = E_DL_VelStep.eRunning) AND iAxis.bError THEN
    bFaultLatch := TRUE;                         // 故障级锁存，仅新启动沿解除
    uErrorId := 16#0004_0230;
    bBusy := FALSE;
    eStep := E_DL_VelStep.eIdle;
END_IF

// 段 7｜速度模式状态机（ENUM + CASE + ELSE 兜底）
CASE eStep OF

    E_DL_VelStep.eIdle:                          // 空闲态：等待启动沿与门禁
        bBusy := FALSE;
        IF rtrigStart.Q THEN
            bFaultLatch := FALSE;                // 新启动沿：锁存码解除路径（R15）
            IF NOT bParamOk THEN
                uErrorId := 16#0004_0106;        // 参数门禁拒绝（信息级）
            ELSIF (iAxis.eState <> E_DL_AxisState.eStandstill)
              AND (iAxis.eState <> E_DL_AxisState.eContinuousMotion) THEN
                uErrorId := 16#0004_0107;        // 非受理态（停止中/故障态）：请求不被受理（信息级）
            ELSE
                fVelEff := fVelocity;            // 目标速度初值 [mm/s]
                IF fVelEff > fVelLim THEN
                    fVelEff := fVelLim;          // 正向超限钳位 [mm/s]
                    uErrorId := 16#0004_0107;    // 信息级：速度钳位提示
                ELSIF fVelEff < -fVelLim THEN
                    fVelEff := -fVelLim;         // 负向超限钳位 [mm/s]
                    uErrorId := 16#0004_0107;    // 信息级：速度钳位提示
                END_IF
                IF (fVelEff <> fVelEff) OR (ABS(fVelEff) > DL_VEL_INF_MAX) THEN
                    fVelEff := 0.0;              // 非有限速度防御归零（0=原地保持，安全侧）
                    uErrorId := 16#0004_0106;    // 信息级：参数门禁拒绝
                END_IF
                IF iAxis.MoveVelocity(fVelEff, fAccEff) THEN
                    fVelSent := fVelEff;         // 记录已发速度，作为改速差值基准 [mm/s]
                    eStep := E_DL_VelStep.eRunning;
                    bBusy := TRUE;
                ELSE
                    bFaultLatch := TRUE;         // 指令被轴拒绝：故障级锁存
                    uErrorId := 16#0004_0230;
                END_IF
            END_IF
        END_IF

    E_DL_VelStep.eRunning:                       // 运行态：电平需求语义 + 动态改速
        bBusy := TRUE;
        IF bCmdStart THEN
            fVelEff := fVelocity;                // 目标速度初值 [mm/s]
            IF fVelEff > fVelLim THEN
                fVelEff := fVelLim;              // 正向超限钳位 [mm/s]
                uErrorId := 16#0004_0107;        // 信息级：速度钳位提示
            ELSIF fVelEff < -fVelLim THEN
                fVelEff := -fVelLim;             // 负向超限钳位 [mm/s]
                uErrorId := 16#0004_0107;        // 信息级：速度钳位提示
            END_IF
            IF (fVelEff <> fVelEff) OR (ABS(fVelEff) > DL_VEL_INF_MAX) THEN
                fVelEff := 0.0;                  // 非有限速度防御归零（安全侧：请求停车速度）
                uErrorId := 16#0004_0106;        // 信息级：参数门禁拒绝
            END_IF
            IF iAxis.eState = E_DL_AxisState.eStandstill THEN
                // 轴已回待机（如限位自动停车）而需求电平仍为真：按电平需求重新发起
                IF iAxis.MoveVelocity(fVelEff, fAccEff) THEN
                    fVelSent := fVelEff;
                ELSE
                    bFaultLatch := TRUE;         // 重发被拒：故障级锁存
                    uErrorId := 16#0004_0230;
                    bBusy := FALSE;
                    eStep := E_DL_VelStep.eIdle;
                END_IF
            ELSIF bDynamicRetarget AND (ABS(fVelEff - fVelSent) > DL_VEL_TGT_TOL) THEN
                // 动态改速：连续运动中差值超容差 → 重发改速（改速而非重启，接口契约语义）
                IF iAxis.eState = E_DL_AxisState.eContinuousMotion THEN
                    IF iAxis.MoveVelocity(fVelEff, fAccEff) THEN
                        fVelSent := fVelEff;     // 更新已发速度基准 [mm/s]
                    ELSE
                        bFaultLatch := TRUE;     // 改速指令被拒：故障级锁存
                        uErrorId := 16#0004_0230;
                        bBusy := FALSE;
                        eStep := E_DL_VelStep.eIdle;
                    END_IF
                ELSE
                    uErrorId := 16#0004_0107;    // 改速请求在非受理态被拒（信息级，瞬态）
                END_IF
            END_IF
        END_IF

    ELSE
        // 非法状态兜底（故障级，沿用族码 0004_0201，复用留档）
        uErrorId := 16#0004_0201;
        bFaultLatch := TRUE;
        bBusy := FALSE;
        eStep := E_DL_VelStep.eIdle;

END_CASE

// 段 8｜状态出口派生（R21：bActive 为轴状态轮询派生式，逐拍重算）
bActive := (iAxis.eState = E_DL_AxisState.eContinuousMotion);
END_FUNCTION_BLOCK

(* ---- FB_DL_BacklashCompensator.st ---- *)
(*
    FB_DL_BacklashCompensator —— 换向背隙补偿
    ------------------------------------------------------------------
    分类      : DL_Motion / Compensation
    前缀      : FB_DL_
    版本      : 1.0.1
    溯源      : T1-6 轴级补偿语义（只借「换向补偿属运动层给定量修正」的分类事实）；
                T2-2 LBP 泵 / 辊「背隙两阶段逼近」组织方式为次源（该组织已被
                RollerGapAdjust 使用）；增量式补偿、EWMA 学习、容差闸与码位 100% 自有；
                clean-room 重写，未复制任何闭源厂商源码，参考实现仅限 MIT/Apache 许可
    平台      : 纯 IEC 61131-3，CODESYS V3.5+ / TwinCAT 3 / InoProShop 通用
    作者      : 道莅代码库 · PLC编程专家（R18）
    ------------------------------------------------------------------
    功能说明  : 指令方向翻转瞬间在给定量上叠加一个方向性补偿量，抵消齿轮 / 丝杠反向
                间隙；并在到位后按实测偏差用 EWMA 自学习背隙估计（现场背隙随磨损变化）；
                与 FB_DL_RollerGapAdjust 的分界是后者为工艺辊缝调整顺控，本件是轴级
                给定量修正，两者不重叠；
                三道闸：负背隙取绝对值（参数习惯差异，不是故障）→ 超上限判故障
                （10 mm 以上补偿会把轴推到撞块）→ 位置非有限即旁路并清方向记忆；
                方向判定带死区，浮点判等全部带容差，杜绝边界来回翻转导致的补偿抖动；
                首拍没有历史方向时绝不补偿，否则轴会凭空跳一下。
    错误码    : 16#0004_01CB 背隙标称值为负已取绝对值 / 学习值被钳位——信息级，不置故障
                16#0004_01CC 预留禁用（信息级，不得挪用）
                16#0004_02DB 背隙标称值超上限（大于 10 mm）——故障级，补偿禁用并旁路输出
                16#0004_02DC 位置快照非有限（NaN / 正负 INF）——故障级，旁路输出并清方向记忆
                16#0004_02DD 预留禁用（故障级，不得挪用）
    码位总账  : 16#0004_01CB 用 / 16#0004_01CC 预留 ｜ 16#0004_02DB 用 / 16#0004_02DC 用 / 16#0004_02DD 预留
    状态机    : 无 CASE，方向由 bPrevDir 一个比特承载，非法状态不可能出现
    采样约定  : fbTrigReset 在本体首部无条件刷新；本件无时间量，补偿结果与任务周期无关，
                自学习按拍迭代，采样越密学习越平滑。
    修订记录  : 2026-11-16 v1.0.0 首次入库（R18）
                2026-11-16 v1.0.1 R18 终审修复：学习率下限常量 DL_BL_MIN_LEARN = 0.001 与引脚声明域
                0.01~0.5 不一致，改为 0.01 与声明对齐（EWMA 仍可双向收敛，无「只置不销」问题）。
                对外引脚零变更。
*)
FUNCTION_BLOCK FB_DL_BacklashCompensator
VAR_INPUT
    bEnable      : BOOL;                       // 使能，FALSE 时输出等于指令（旁路）/ enable, FALSE passes the command through
    bReset       : BOOL;                       // 上升沿清方向记忆与学习值 / rising edge clears the direction memory and the learned value
    fCmdPosition : REAL := 0.0;                // 指令位置，来自插补或定位 [mm] / commanded position from the interpolator or the positioner [mm]
    fActPosition : REAL := 0.0;                // 实际位置反馈，自学习用 [mm] / actual position feedback used for learning [mm]
    fBacklash    : REAL := 0.10;               // 背隙标称值 [mm]，范围 0.0~10.0 / nominal backlash [mm], range 0.0~10.0
    bAutoLearn   : BOOL := FALSE;              // TRUE 时按到位偏差 EWMA 更新背隙 / TRUE updates the backlash from the positioning deviation by EWMA
    fLearnTol    : REAL := 0.10;               // 学习容差，到位偏差超此值不采信 [mm] / learning tolerance, deviations above it are rejected [mm]
    fLearnGain   : REAL := 0.1;                // EWMA 学习率 [无量纲]，范围 0.01~0.5 / EWMA learning rate [dimensionless], range 0.01~0.5
END_VAR
VAR_OUTPUT
    fOutPosition : REAL;                       // 补偿后位置给定 [mm] / compensated position setpoint [mm]
    bDirPositive : BOOL;                       // 当前指令方向，TRUE 为正向 / current command direction, TRUE is positive
    fApplied     : REAL;                       // 本拍叠加的补偿量（带符号）[mm] / compensation applied this cycle with its sign [mm]
    fBacklashEst : REAL;                       // 当前背隙估计（学习值）[mm] / current backlash estimate [mm]
    bLearnActive : BOOL;                       // 本次自学习被采信 / this cycle learning was accepted
    eErr         : UDINT;                      // 错误码，0=正常 / error id, 0=ok
    bError       : BOOL;                       // 故障标志，eErr 为故障级时 TRUE / error flag, TRUE on fault-level eErr
END_VAR
VAR
    fbTrigReset : R_TRIG;                      // 复位沿检测实例，本体首部无条件刷新 / reset edge instance, refreshed unconditionally
    bPrevDir    : BOOL;                        // 上一拍方向，TRUE 正向 / previous cycle direction, TRUE is positive
    bDirInit    : BOOL := FALSE;               // 方向记忆已初始化标志，初值 FALSE / direction memory initialised flag, initial FALSE
    bDirCur     : BOOL;                        // 本拍方向判定结果 / current cycle direction
    bReversed   : BOOL;                        // 方向翻转标志 / direction reversal flag
    bInit       : BOOL := FALSE;               // 首扫标志，初值 FALSE，判据 NOT bInit / first-scan flag, initial FALSE, tested with NOT
    fEst        : REAL;                        // 背隙估计（EWMA 值）[mm] / backlash estimate produced by EWMA [mm]
    fDev        : REAL;                        // 到位偏差，实际减指令 [mm] / positioning deviation, actual minus command [mm]
    fPrevCmd    : REAL;                        // 上一拍指令位置，方向判定用 [mm] / previous commanded position used by the direction check [mm]
    fBlEff      : REAL;                        // 生效背隙标称值，取绝对值后 [mm] / effective nominal backlash after the absolute value [mm]
    fGainEff    : REAL;                        // 生效学习率，钳位后 [无量纲] / effective learning rate after clamping [dimensionless]
    fAppliedInt : REAL;                        // 补偿量中间量 [mm] / compensation intermediate [mm]
    fClamped    : REAL;                        // 钳位中间量 [mm] / clamping intermediate [mm]
    bNonFin     : BOOL;                        // 位置非有限判定标志 / position non-finite flag
END_VAR
VAR CONSTANT
    DL_BL_MAX        : REAL := 10.0;           // 背隙上限 [mm] / backlash upper bound [mm]
    DL_BL_MIN_LEARN  : REAL := 0.01;           // 学习率下限 [无量纲]，与引脚声明域 0.01~0.5 一致 / learning rate lower bound [dimensionless], aligned with the documented 0.01~0.5 pin range
    DL_BL_GAIN_MAX   : REAL := 0.5;            // 学习率上限 [无量纲] / learning rate upper bound [dimensionless]
    DL_BL_INF_GUARD  : REAL := 4.0E38;         // 非有限幅值判定阈值 [mm] / non-finite magnitude guard [mm]
    DL_FLOAT_EPS     : REAL := 1.0E-6;         // 浮点判等容差 [mm] / float equality tolerance [mm]
    DL_BL_ZERO       : REAL := 0.0;            // 零值常量，避免裸字面量 [无量纲] / zero constant, avoids a bare literal [dimensionless]
    DL_BL_ONE        : REAL := 1.0;            // 一值常量，用于符号判定 / one constant used by the sign check [dimensionless]
END_VAR

// 段 1｜边沿实例无条件周期刷新（红线：严禁放入条件分支）/ segment 1, unconditional edge refresh
fbTrigReset(CLK := bReset);

// 段 2｜输出与错误状态预置 / segment 2, preset outputs and error status
eErr := 0;                                     // 预置无错误 / preset no error
bError := FALSE;                               // 预置无故障 / preset no fault
bLearnActive := FALSE;                         // 预置本次不采信学习 / preset learning not accepted
fApplied := DL_BL_ZERO;                        // 补偿量先清零 / clear the applied compensation
bReversed := FALSE;                            // 翻转标志先清 / clear the reversal flag

// 段 3｜首扫初始化（初值 FALSE，判据 NOT bInit）/ segment 3, first-scan initialisation
IF NOT bInit THEN
    fEst := MIN(MAX(ABS(fBacklash), DL_BL_ZERO), DL_BL_MAX); // 初值取标称背隙绝对值，双侧钳位 / initialise from the absolute nominal backlash, clamped both sides
    fPrevCmd := DL_BL_ZERO;                    // 指令记忆清零 / clear the command memory
    bDirInit := FALSE;                         // 方向记忆未初始化 / the direction memory is not initialised yet
    bInit := TRUE;                             // 首扫只做一次 / first scan runs once only
END_IF

// 段 4｜使能闸：旁路输出，不补偿 / segment 4, enable gate passes the command through
IF NOT bEnable THEN
    fOutPosition := fCmdPosition;              // 输出等于指令 / output equals the command
    fBacklashEst := fEst;                      // 估计值照常回读 / the estimate stays readable
    RETURN;                                    // 失能即出口 / disabled is the exit
END_IF

// 段 5｜背隙标称值闸：负值取绝对值（参数习惯），超上限判故障 / segment 5, nominal backlash gate
fBlEff := ABS(fBacklash);                      // 负背隙取绝对值 / take the absolute value of a negative backlash
IF fBacklash < DL_BL_ZERO THEN
    eErr := 16#0004_01CB;                      // 取绝对值提示（信息级不置故障）/ absolute value hint, info level never raises a fault
END_IF
IF fBlEff > DL_BL_MAX THEN
    eErr := 16#0004_02DB;                      // 背隙超上限故障码 / backlash above the cap fault id
    bError := TRUE;                            // 置故障标志 / raise the error flag
    fOutPosition := fCmdPosition;              // 补偿禁用，旁路输出 / compensation disabled, pass the command through
    fBacklashEst := fEst;                      // 估计值回读 / the estimate stays readable
    RETURN;                                    // 故障级提前返回 / early return on fault
END_IF

// 段 6｜位置非有限闸：旁路输出并清方向记忆 / segment 6, non-finite position gate
bNonFin := (fCmdPosition <> fCmdPosition)
        OR (fCmdPosition > DL_BL_INF_GUARD) OR (fCmdPosition < -DL_BL_INF_GUARD)
        OR (fActPosition <> fActPosition)
        OR (fActPosition > DL_BL_INF_GUARD) OR (fActPosition < -DL_BL_INF_GUARD); // 双位置同口径检查 / both positions checked the same way
IF bNonFin THEN
    eErr := 16#0004_02DC;                      // 位置非有限故障码 / non-finite position fault id
    bError := TRUE;                            // 置故障标志 / raise the error flag
    fOutPosition := fCmdPosition;              // 旁路输出 / pass the command through
    fBacklashEst := fEst;                      // 估计值回读 / the estimate stays readable
    bDirInit := FALSE;                         // 清方向记忆，防下一拍凭空跳一下 / clear the direction memory so the next cycle cannot jump
    RETURN;                                    // 故障级提前返回 / early return on fault
END_IF

// 段 7｜首拍无历史方向：不补偿，只登记方向 / segment 7, no compensation without a historical direction
IF NOT bDirInit THEN
    fPrevCmd := fCmdPosition;                  // 登记指令位置 / register the commanded position
    bPrevDir := TRUE;                          // 默认按正向登记 / register the positive direction by default
    bDirInit := TRUE;                          // 方向记忆就绪 / the direction memory is ready
    bDirPositive := TRUE;                      // 对外方向 / publish the direction
    fOutPosition := fCmdPosition;              // 首拍不补偿 / no compensation on the first cycle
    fBacklashEst := fEst;                      // 估计值回读 / the estimate stays readable
    RETURN;                                    // 本拍结束 / the cycle ends here
END_IF

// 段 8｜方向判定：带死区，浮点判等全部带容差，死区内保持上一方向 / segment 8, direction detection with a dead band
IF fCmdPosition > (fPrevCmd + DL_FLOAT_EPS) THEN
    bDirCur := TRUE;                           // 越过死区向上，判正向 / above the dead band, positive
ELSIF fCmdPosition < (fPrevCmd - DL_FLOAT_EPS) THEN
    bDirCur := FALSE;                          // 越过死区向下，判负向 / below the dead band, negative
ELSE
    bDirCur := bPrevDir;                       // 死区内保持上一方向，防抖动翻转 / inside the dead band keep the previous direction against chatter
END_IF
bReversed := (bDirCur <> bPrevDir);            // 方向翻转判定 / reversal detection
bDirPositive := bDirCur;                       // 对外方向 / publish the direction

// 段 9｜复位沿：清方向记忆与学习值（优先于补偿）/ segment 9, reset clears the direction memory and the learned value
IF fbTrigReset.Q THEN
    fEst := MIN(MAX(fBlEff, DL_BL_ZERO), DL_BL_MAX); // 学习值回到标称 / the learned value returns to the nominal
    fPrevCmd := fCmdPosition;                  // 指令记忆复位 / reset the command memory
    bDirInit := FALSE;                         // 方向记忆清空 / clear the direction memory
    bReversed := FALSE;                        // 本拍不判翻转 / no reversal on the reset cycle
    fOutPosition := fCmdPosition;              // 复位拍不补偿 / no compensation on the reset cycle
    fBacklashEst := fEst;                      // 估计值回读 / the estimate stays readable
    RETURN;                                    // 复位即出口 / reset is the exit
END_IF

// 段 10｜EWMA 自学习：仅在非翻转拍、偏差在容差内且非零时采信 / segment 10, EWMA learning accepted only off the reversal cycle
fGainEff := MIN(MAX(fLearnGain, DL_BL_MIN_LEARN), DL_BL_GAIN_MAX); // 学习率双侧钳位 / clamp the learning rate both sides
IF (ABS(fLearnGain - fGainEff) > DL_FLOAT_EPS) THEN
    eErr := 16#0004_01CB;                      // 学习率钳位提示（信息级不置故障）/ learning rate clamp hint, info level never raises a fault
END_IF
IF bAutoLearn AND (NOT bReversed) THEN
    fDev := fActPosition - fCmdPosition;       // 到位偏差 / positioning deviation
    IF (ABS(fDev) <= fLearnTol) AND (ABS(fDev) > DL_FLOAT_EPS) THEN
        fEst := fEst + fGainEff * (ABS(fDev) - fEst); // 一阶 EWMA 逼近偏差绝对值 / first order EWMA towards the absolute deviation
        fClamped := MIN(MAX(fEst, DL_BL_ZERO), DL_BL_MAX); // 学习值双侧钳位 / clamp the learned value both sides
        IF ABS(fClamped - fEst) > DL_FLOAT_EPS THEN
            eErr := 16#0004_01CB;              // 学习值钳位提示（信息级不置故障）/ learned value clamp hint, info level never raises a fault
        END_IF
        fEst := fClamped;                      // 落盘钳位值 / commit the clamped value
        bLearnActive := TRUE;                  // 本次学习被采信 / this cycle learning is accepted
    END_IF
END_IF

// 段 11｜补偿量与输出：幅值不超过背隙上限，方向翻转即换符号，恒定而非逐拍累加 / segment 11, compensation and output
IF bDirCur THEN
    fAppliedInt := fEst;                       // 正向运动叠加正补偿 / a positive move carries a positive compensation
ELSE
    fAppliedInt := -fEst;                      // 负向运动叠加负补偿 / a negative move carries a negative compensation
END_IF
IF ABS(fAppliedInt) > DL_BL_MAX THEN
    IF fAppliedInt >= DL_BL_ZERO THEN
        fAppliedInt := DL_BL_MAX;              // 正向幅值兜底钳位 / positive magnitude fallback clamp
    ELSE
        fAppliedInt := -DL_BL_MAX;             // 负向幅值兜底钳位 / negative magnitude fallback clamp
    END_IF
END_IF
fApplied := fAppliedInt;                       // 对外补偿量 / publish the compensation
fOutPosition := fCmdPosition + fAppliedInt;    // 补偿后给定 / compensated setpoint
fBacklashEst := fEst;                          // 对外背隙估计 / publish the backlash estimate

// 段 12｜方向记忆推进 / segment 12, advance the direction memory
fPrevCmd := fCmdPosition;                      // 记录本拍指令 / remember this cycle command
bPrevDir := bDirCur;                           // 记录本拍方向 / remember this cycle direction
END_FUNCTION_BLOCK

(* ---- FB_DL_BagFeedDancerSync.st ---- *)
//==============================================================================
// 功能块：FB_DL_BagFeedDancerSync ｜ 中文名称：制袋供膜摆辊同步（复杂度 H）
// 所属子库：DL_Motion ｜ 版本：v1.0.1 ｜ 兼容：CODESYS V3.5+ / TwinCAT 3 / 汇川 InoProShop
// 功能描述：制袋机供膜摆辊同步——供膜速度给定 = 线速前馈 + 摆辊位置 PI
//           修正；摆辊信号不可信时前馈直通、PI 冻结（域外行为显式化）；
//           输出触顶积分冻结（抗饱和）；停链且摆辊持续偏离中位判张力故障。
//           【拓扑语义假设（R23 终审留档，符号判定的前提）】供膜单元位于
//           摆辊环下游（自环内抽膜、与线速同步），摆辊位置偏大 = 环内膜存
//           量过多 → PI 正向修正加快抽膜耗环（负反馈收敛）。若调用方拓扑
//           相反（供膜自环上游推膜），须将 fFeedKp / fFeedKi 反号接入或
//           另行适配，本件不自动判向。
// 开源溯源 (Origin)：道莅原创实现（参考包装制袋机摆辊同步工程惯例 分类与参数域）
// 单位表：摆辊位置[%]（50 = 中位）/ 线速与供膜速度[mm/s] / 增益[（mm/s）/%]
//         与[（mm/s）/(%·拍)] / 速度上限[mm/s] / 计时[ms]
// 错误码表：16#0004_01E1 信息级（摆辊域外/非有限不可信，或线速负值已钳
//           0——共码，不置 bError）/ 16#0004_01E2 预留禁用（不得挪用）/
//           16#0004_02FC 故障级（供膜速度上限组态非法 <= 0，置 bError）/
//           16#0004_02FD 故障级（张力疑似故障：线速 0 且摆辊持续偏离中位
//           超窗，断膜/卡膜疑似，置 bError）/ 16#0004_02FE 故障级兜底
//           （置 bError）
// 状态机：N/A（PI 修正 + 阈值判窗为电平逻辑，无相位状态机）
// 边界行为：① 摆辊位置域外（0~100 外）或非有限 → bDancerOk := FALSE +
//           前馈直通（PI 冻结，积分保持）+ 信息 01E1（R11 NtcTempScan 同
//           口径）；② PI 抗饱和：输出触顶（0 或上限）时积分冻结；③
//           fLineSpeedMmS < 0 → 钳 0 + 信息 01E1 复用（R90）；④
//           fFeedMaxMmS <= 0 → 故障 02FC；⑤ 线速为 0 且摆辊持续偏离中位
//           > tIdleOffTol → bTensionFault := TRUE + 故障 02FD；⑥ 积分增益
//           按拍积分（无周期引脚），有效量纲 [（mm/s）/(%·拍)]，头注释
//           单位表留档此口径。
// 依赖收窄 (R11 留档③)：Motion 不得跨库调用前馈补偿件（FeedforwardComp
//           等均为他库），前馈律（fFeedSp := fLineSpeed + PI 修正）在本件
//           内联实现，改动任一侧须复核另一侧。
// 修订历史：v1.0.0 2026-11-17 首版（R23 派单 · ROADMAP 包装 P1 §377）
//           v1.0.1 2026-11-17 R23 终审补档（逻辑零改动）：头注释补拓扑
//           语义假设声明——PI 符号经推演在「抽膜」拓扑下为负反馈正确，
//           但原版未留档流向假设，反拓扑接入会翻转为正反馈发散。
//==============================================================================

FUNCTION_BLOCK FB_DL_BagFeedDancerSync
VAR_INPUT
    fDancerPosPct : LREAL;                  // 摆辊位置 [百分数]，50 = 中位，有效域 0..100 / Dancer position [percent], 50 = mid
    fLineSpeedMmS : LREAL;                  // 线速前馈源 [毫米/秒] / Line speed feedforward source [mm/s]
    fFeedKp       : LREAL := 1.5;           // 摆辊 PI 比例增益 [（毫米/秒）/%] / Dancer PI proportional gain [(mm/s)/%]
    fFeedKi       : LREAL := 0.2;           // 摆辊 PI 积分增益 [（毫米/秒）/(%·拍)]，按拍积分 / Dancer PI integral gain per scan
    fFeedMaxMmS   : LREAL := 500.0;         // 供膜速度上限 [毫米/秒]，须 > 0 / Feed speed ceiling [mm/s], must be > 0
    bEnable       : BOOL;                   // 同步使能 [—] / Sync enable
    bReset        : BOOL;                   // 故障复位 [—]，清除张力故障锁存 / Fault reset, clears the tension latch
END_VAR
VAR_OUTPUT
    fFeedSpMmS    : LREAL;                  // 供膜速度给定 [毫米/秒] = 前馈 + PI 修正 / Feed speed setpoint [mm/s] = feedforward plus PI trim
    bDancerOk     : BOOL;                   // 摆辊信号可信 [—] / Dancer signal trustworthy
    bTensionFault : BOOL;                   // 张力疑似故障 [—] / Tension suspected fault
    eErr          : UDINT;                  // 错误码，0 = 无错 / Error code, 0 = no error
    bError        : BOOL;                   // 故障级标志，仅故障级错误置位 / Fault-class flag, set only on fault-level codes
    bValid        : BOOL;                   // 输出可用标志 / Outputs usable flag
END_VAR
VAR
    fbIdleOff     : TON;                    // 停链偏离中位判窗，段 6 无条件刷新 [ms] / Idle off-mid window
    _fPosEff      : LREAL;                  // 生效摆辊位置 [百分数] / Effective dancer position [percent]
    _fLineEff     : LREAL;                  // 钳位后的生效线速 [毫米/秒] / Effective clamped line speed [mm/s]
    _fErr         : LREAL;                  // 摆辊位置偏差 [百分数] / Dancer position error [percent]
    _fPITrim      : LREAL;                  // PI 修正量 [毫米/秒] / PI trim [mm/s]
    _fIntAcc      : LREAL;                  // 积分累加器 [毫米/秒] / Integral accumulator [mm/s]
    _bInit        : BOOL := FALSE;          // 首扫标志，初值 FALSE 取非判定 / First-scan flag, tested negated
    _bDancerBad   : BOOL;                   // 摆辊不可信当拍标志 / Dancer-untrustworthy flag of this scan
    _bLineClamp   : BOOL;                   // 线速钳位当拍标志 / Line clamp flag of this scan
    _bCfgBad      : BOOL;                   // 速度上限组态非法锁存 / Illegal ceiling latch
    _bTensionLatch: BOOL;                   // 张力故障锁存（bReset 清除） / Tension fault latch, cleared by bReset
    _bIllegal     : BOOL;                   // 非法状态标志 / Illegal state flag
END_VAR
VAR CONSTANT
    DL_BF_POS_MIN : LREAL := 0.0;           // 摆辊位置域下限 [百分数] / Dancer position domain floor [percent]
    DL_BF_POS_MAX : LREAL := 100.0;         // 摆辊位置域上限 [百分数] / Dancer position domain ceiling [percent]
    DL_BF_MID     : LREAL := 50.0;          // 摆辊中位 [百分数] / Dancer mid position [percent]
    DL_BF_IDLE_TOL: LREAL := 10.0;          // 停链偏离中位容差 [百分数] / Idle off-mid tolerance [percent]
    DL_BF_IDLE_WIN: TIME  := T#5S;          // 停链偏离判窗 [ms] / Idle off-mid window [ms]
    DL_BF_INF     : LREAL := 1.7976931348623157E308; // LREAL 幅值上限 / LREAL magnitude ceiling
    DL_BF_EPS     : LREAL := 1.0E-6;        // 浮点判零容差 [毫米/秒] / Float zero tolerance [mm/s]
END_VAR

(*------------------------------------------------------------------------------
 * 段 1｜每拍预置：输出先算后出，单拍标志预清零
 *      Outputs computed per scan, one-shot flags pre-cleared
 *-----------------------------------------------------------------------------*)
fFeedSpMmS  := 0.0;                         // 供膜给定预置零 / Feed setpoint preset zero
bDancerOk   := FALSE;                       // 可信标志预置 FALSE / Trustworthy preset FALSE
bTensionFault := FALSE;                     // 张力故障每拍重算 / Tension fault recomputed
eErr        := 16#0000_0000;                // 错误码每拍重算 / Error code recomputed
bError      := FALSE;                       // 故障标志每拍重算 / Fault flag recomputed
bValid      := FALSE;                       // 可用标志每拍重算 / Usable flag recomputed
_bDancerBad := FALSE;                       // 摆辊标志预清零 / Dancer flag pre-cleared
_bLineClamp := FALSE;                       // 线速钳位预清零 / Line clamp pre-cleared
_bIllegal   := FALSE;                       // 非法状态预清零 / Illegal flag pre-cleared

(*------------------------------------------------------------------------------
 * 段 2｜首扫初始化
 *      First-scan initialisation
 *-----------------------------------------------------------------------------*)
IF NOT _bInit THEN
    _fIntAcc  := 0.0;                       // 积分累加器清零 / Integral accumulator cleared
    _bCfgBad  := FALSE;                     // 组态锁存清零 / Config latch cleared
    _bTensionLatch := FALSE;                // 张力锁存清零 / Tension latch cleared
    _bInit    := TRUE;                      // 首扫只做一次 / The first scan runs once
END_IF

(*------------------------------------------------------------------------------
 * 段 3｜组态与输入防御闸（速度上限 <= 0 → 02FC；摆辊/线速非有限 → 不可信）
 *      Configuration and input defense gates
 *-----------------------------------------------------------------------------*)
IF (fFeedMaxMmS <> fFeedMaxMmS) OR (ABS(fFeedMaxMmS) > DL_BF_INF) OR (fFeedMaxMmS <= 0.0) THEN
    _bCfgBad := TRUE;                       // 速度上限组态非法锁存 / Illegal ceiling latched
END_IF
IF (fDancerPosPct <> fDancerPosPct) OR (ABS(fDancerPosPct) > DL_BF_INF)
   OR (fLineSpeedMmS <> fLineSpeedMmS) OR (ABS(fLineSpeedMmS) > DL_BF_INF)
   OR (fFeedKp <> fFeedKp) OR (ABS(fFeedKp) > DL_BF_INF)
   OR (fFeedKi <> fFeedKi) OR (ABS(fFeedKi) > DL_BF_INF) THEN
    _bDancerBad := TRUE;                    // 任一输入非有限：摆辊判不可信（R79） / Any non-finite input, dancer untrustworthy
END_IF

(*------------------------------------------------------------------------------
 * 段 4｜摆辊域外与线速钳位（域外行为显式化，信息级共码 01E1，R90）
 *      Out-of-domain handling with a shared info code per R90
 *-----------------------------------------------------------------------------*)
IF (NOT _bDancerBad) AND ((fDancerPosPct < DL_BF_POS_MIN) OR (fDancerPosPct > DL_BF_POS_MAX)) THEN
    _bDancerBad := TRUE;                    // 摆辊域外：不可信（前馈直通） / Dancer out of domain, untrustworthy
END_IF
IF fLineSpeedMmS < 0.0 THEN
    _fLineEff := 0.0;                       // 负线速钳 0（物理下界） / Negative line speed clamped to zero
    _bLineClamp := TRUE;                    // 钳位声明 / Clamp declared
ELSE
    _fLineEff := fLineSpeedMmS;             // 合法线速原值生效 / Valid line speed applied as-is
END_IF

(*------------------------------------------------------------------------------
 * 段 5｜PI 修正与前馈合成（可信时积分推进，不可信/触顶冻结——抗饱和）
 *      PI trim and feedforward synthesis with anti-windup freezing
 *-----------------------------------------------------------------------------*)
IF bEnable AND (NOT _bCfgBad) AND (NOT _bDancerBad) THEN
    bDancerOk := TRUE;                      // 摆辊可信 / Dancer trustworthy
    _fPosEff := fDancerPosPct;              // 生效位置原值 / Effective position as-is
    _fErr := _fPosEff - DL_BF_MID;          // 位置偏差 [百分数]，偏大 = 膜存量过多 / Position error, high means excess film stored
    _fPITrim := fFeedKp * _fErr + _fIntAcc; // PI 修正量 [毫米/秒] / PI trim [mm/s]
    fFeedSpMmS := _fLineEff + _fPITrim;     // 供膜给定 = 前馈 + 修正 / Feed setpoint = feedforward plus trim
    IF fFeedSpMmS < 0.0 THEN
        fFeedSpMmS := 0.0;                  // 下限钳 0（反向不倒转） / Lower clamp, no reverse
        (* 输出触下限：积分冻结（抗饱和） / Saturated at the floor, integral frozen *)
    ELSIF fFeedSpMmS > fFeedMaxMmS THEN
        fFeedSpMmS := fFeedMaxMmS;          // 上限钳位 / Ceiling clamp
        (* 输出触上限：积分冻结（抗饱和） / Saturated at the ceiling, integral frozen *)
    ELSE
        _fIntAcc := _fIntAcc + fFeedKi * _fErr; // 未触顶：积分推进（按拍积分） / Not saturated, integral advances per scan
    END_IF
ELSE
    (* 摆辊不可信：前馈直通（PI 冻结，积分保持不推进） / Untrustworthy, feedforward passthrough, integral held *)
    fFeedSpMmS := _fLineEff;                // 前馈直通 / Feedforward passthrough
    IF fFeedSpMmS > fFeedMaxMmS THEN
        fFeedSpMmS := fFeedMaxMmS;          // 直通仍受上限约束 / Passthrough still ceiling-clamped
    END_IF
    IF fFeedSpMmS < 0.0 THEN
        fFeedSpMmS := 0.0;                  // 直通仍受下限约束 / Passthrough still floor-clamped
    END_IF
    IF _bDancerBad OR _bLineClamp THEN
        bDancerOk := FALSE;                 // 不可信声明出口 / Untrustworthy declared
    END_IF
END_IF

(*------------------------------------------------------------------------------
 * 段 6｜停链偏离判窗无条件刷新（R40：CASE 之外每拍必调）
 *      Idle off-mid window refreshed unconditionally per R40
 *-----------------------------------------------------------------------------*)
fbIdleOff(IN := bEnable AND (NOT _bCfgBad) AND (NOT _bDancerBad)
              AND (_fLineEff <= DL_BF_EPS)
              AND (ABS(fDancerPosPct - DL_BF_MID) > DL_BF_IDLE_TOL), PT := DL_BF_IDLE_WIN); // 停链偏离中位判窗 / Idle off-mid window
IF fbIdleOff.Q THEN
    _bTensionLatch := TRUE;                 // 张力故障锁存（断膜/卡膜疑似） / Tension fault latched
END_IF
IF bReset THEN
    _bTensionLatch := FALSE;                // 复位清张力锁存 / Reset clears the tension latch
END_IF
bTensionFault := _bTensionLatch;            // 张力故障出口 / Tension fault outlet

(*------------------------------------------------------------------------------
 * 段 7｜码位出口
 *      Code outlet
 *-----------------------------------------------------------------------------*)
IF _bCfgBad THEN
    eErr   := 16#0004_02FC;                 // 故障级：速度上限组态非法 / Fault: illegal speed ceiling
    bError := TRUE;                         // 置故障标志（R45 配对） / Raise the fault flag
    bValid := FALSE;                        // 输出不可用 / Outputs unusable
ELSIF _bTensionLatch THEN
    eErr   := 16#0004_02FD;                 // 故障级：张力疑似故障 / Fault: tension suspected
    bError := TRUE;                         // 置故障标志 / Raise the fault flag
    bValid := TRUE;                         // 判定结果本身可用 / The verdict itself is usable
ELSIF _bDancerBad OR _bLineClamp THEN
    eErr := 16#0004_01E1;                   // 信息级：摆辊/线速已钳位或不可信（共码，R90） / Info: clamped or untrustworthy, shared code
    bValid := TRUE;                         // 前馈直通结果可用（降级口径） / Passthrough result usable
ELSE
    bValid := bEnable;                      // 使能且正常：输出可用 / Outputs usable when enabled
END_IF
END_FUNCTION_BLOCK

(* ---- FB_DL_BrakeReleaseInterlock.st ---- *)
(*
    FB_DL_BrakeReleaseInterlock —— 伺服抱闸释放互锁
    ------------------------------------------------------------------
    分类      : DL_Motion / AxisSafety
    前缀      : FB_DL_
    版本      : 1.0.0
    溯源      : clean-room 自有实现；仅借鉴「先确认力矩再放闸」的公开工程常识语义，
                未复制任何闭源厂商源码，码位 100% 自有
    平台      : 纯 IEC 61131-3，CODESYS V3.5+ / TwinCAT 3 / InoProShop / Machine Expert 通用
    作者      : 道莅代码库 · PLC编程专家（R76 冲刺批 C3 · #1）
    ------------------------------------------------------------------
    功能说明  : 伺服抱闸「释放侧互锁」唯一时序属主件：伺服使能建立 → 力矩到达确认
                （fTorque < fReleaseTh 持续 tTorqueQual）→ 发抱闸释放输出 →
                闸位反馈确认（bBrakeReleased）→ 就绪（bReady）。
                边界：只产出抱闸释放命令与就绪标志，不发运动指令、不直控伺服使能；
                与 FB_DL_AxisBrakeSeq（上/断电两条全序）差异化：本件聚焦
                「释放互锁单序 + 运行中失使能即时回闸」。
    序列      : eIdle --bServoEnabled--> eTorqueQual --fbTorqueQual.Q--> eReleasing
                --bBrakeReleased--> eReady；
                eReady --bServoEnabled丢失--> eClosing（立即撤输出重上闸）
                --反馈闭合或 tCloseWait--> eIdle；
                eReleasing --tReleaseTimeout--> eFault（撤输出回退，弹簧闸抱死为安全侧）；
                任意态 --参数/采样非法--> eFault。
    错误码    : 16#0005_1D00 力矩确认超时（tTorqueQual 内未持续低于阈值）——故障级，撤输出回退
                16#0005_1D01 抱闸释放反馈超 tReleaseTimeout——故障级，撤输出回退
                16#0005_1D02 就绪态伺服使能丢失，已立即重新上闸——信息级，eClosing 期间持续发布
                16#0005_1D03 时序中途使能丢失，回退重新上闸——信息级，eClosing 期间持续发布
                16#0005_1D04 力矩采样非有限（NaN 用 f<>f、±Inf 用 (f-f)<>(f-f)）——故障级
                16#0005_1D05 参数非法（阈值非正 / 任一时间为零）——故障级
                16#0005_1D06 就绪态释放反馈意外跌落（抱闸非受控闭合）——故障级
                16#0005_1D07 CASE 落 ELSE 兜底——故障级
    码位总账  : 16#0005_1D00..1D07 全部定义并使用，无空悬码位
    状态机    : E_DL_BrakeRelState（eIdle / eTorqueQual / eReleasing / eReady / eClosing
                / eFault），CASE 含 ELSE 兜底：落 ELSE 置 16#0005_1D07、撤输出回 eFault。
                故障码锁存至复位沿：bReset 上升沿且 bServoEnabled=FALSE 时方可复位
                （带使能复位会立即重新放闸，禁止）；信息级码不置 bError、随相发布。
    定时器    : 三只 TON + 一只 R_TRIG 在本体段 1 无条件周期刷新（R7），绝不放入 CASE/IF；
                相转出靠状态条件失配自然断输入，无跨相复用实例。
    防御口径  : 浮点比较一律阈值/容差，禁 =/<>；本件无除法运算；非有限判定按
                NaN f<>f、±Inf (f-f)<>(f-f) 双判，不近似阈值。
    修订记录  : 2026-11-23 v1.0.0 首次入库（R76 冲刺批 C3 · #1）
*)
TYPE E_DL_BrakeRelState :
(
    eIdle       := 0,   // 待机，释放命令失电，等伺服使能建立 / idle, release command off, waiting for the servo enable
    eTorqueQual := 10,  // 力矩确认中，fTorque 持续低于阈值计时 / torque qualifying, timing while torque stays under threshold
    eReleasing  := 20,  // 已发释放命令，等闸位反馈确认 / release command asserted, waiting for brake feedback
    eReady      := 30,  // 释放互锁就绪，抱闸已开且使能在 / interlock ready, brake open and enable present
    eClosing    := 40,  // 回闸中，命令已撤，等反馈闭合或时间兜底 / re-closing, command off, waiting for closed feedback or the fallback time
    eFault      := 50   // 故障，撤输出回退，故障码锁存至复位沿 / fault, outputs rolled back, code latched until reset edge
);
END_TYPE

FUNCTION_BLOCK FB_DL_BrakeReleaseInterlock
VAR_INPUT
    bServoEnabled    : BOOL;              // 伺服使能状态，TRUE = 使能已建立 / servo enable status, TRUE = enable established
    fTorque          : REAL;              // 伺服当前力矩 [Nm]，参与确认判定 / servo torque [Nm], used by the qualification test
    fReleaseTh       : REAL := 5.0;       // 力矩确认阈值 [Nm]，必须大于 0 / torque qualification threshold [Nm], must exceed zero
    tTorqueQual      : TIME := T#300MS;   // 力矩确认持续时间 [ms]，必须大于 0 / torque qualification dwell [ms], must exceed zero
    bBrakeReleased   : BOOL;              // 抱闸释放到位反馈，TRUE = 已完全释放 / brake released feedback, TRUE = fully released
    tReleaseTimeout  : TIME := T#3S;      // 释放反馈超时 [ms]，必须大于 0 / release feedback timeout [ms], must exceed zero
    tCloseWait       : TIME := T#500MS;   // 回闸兜底等待 [ms]，反馈闭合可提前退出 / re-close fallback wait [ms], closed feedback exits earlier
    bReset           : BOOL;              // 故障复位请求，上升沿生效且须无使能 / fault reset request, edge-active and requires no enable
END_VAR
VAR_OUTPUT
    bBrakeReleaseCmd : BOOL;              // 抱闸释放命令输出，仅 eReleasing/eReady 置位 / brake release command, asserted in eReleasing/eReady only
    bReady           : BOOL;              // 释放互锁就绪标志 / release interlock ready flag
    eState           : E_DL_BrakeRelState; // 当前状态镜像输出 / current state mirror output
    nErrCode         : UDINT;             // 错误码，0 = 无错；信息级随相发布、故障级锁存回放 / error code, 0 = none; info codes published per phase, fault codes latched
    bError           : BOOL;              // 故障级标志，仅故障级码置位 / fault-class flag, raised only by fault-class codes
    bValid           : BOOL;              // 输出可用标志，= NOT bError / outputs valid flag, equals NOT bError
END_VAR
VAR
    fbTorqueQual     : TON;               // 力矩确认定时器，仅 eTorqueQual 使用 / torque qualification timer, eTorqueQual only
    fbReleaseTo      : TON;               // 释放反馈超时定时器，仅 eReleasing 使用 / release feedback timeout timer, eReleasing only
    fbCloseWait      : TON;               // 回闸兜底定时器，仅 eClosing 使用 / re-close fallback timer, eClosing only
    rtReset          : R_TRIG;            // 复位上升沿检测 / reset rising-edge detector
    _eState          : E_DL_BrakeRelState; // 当前状态 / current state
    _uErrLatch       : UDINT;             // 故障码锁存副本，故障态每拍回放 / latched fault code republished inside the fault state
    _bGateOk         : BOOL;              // 参数与采样门禁结果 / parameter and sample gate result
    _bLostInReady    : BOOL;              // TRUE = 就绪态丢使能（1D02），FALSE = 中途丢（1D03）/ TRUE = enable lost in eReady (1D02), FALSE = lost mid-sequence (1D03)
END_VAR
VAR CONSTANT
    DL_BRI_ZERO : REAL := 0.0;            // 零值常量，避免裸字面量 [Nm] / zero constant avoiding a bare literal [Nm]
    DL_BRI_T_ZERO : TIME := T#0S;         // 零时间常量，参数门禁用 / zero time constant for the parameter gate
END_VAR

// 段 1｜定时器与边缘检测无条件周期刷新（R7：严禁放入 IF / CASE，实例无跨相复用）
// segment 1, timers and edge detectors refreshed unconditionally, never inside IF/CASE, no cross-phase reuse
fbTorqueQual(IN := (_eState = E_DL_BrakeRelState.eTorqueQual) AND _bGateOk, PT := tTorqueQual);
fbReleaseTo(IN := (_eState = E_DL_BrakeRelState.eReleasing), PT := tReleaseTimeout);
fbCloseWait(IN := (_eState = E_DL_BrakeRelState.eClosing), PT := tCloseWait);
rtReset(CLK := bReset);

// 段 2｜输出与错误状态预置；故障态从锁存副本回放（故障码锁存至复位沿，不被预置冲掉）
// segment 2, preset outputs and error status; the fault state replays from the latch so the preset cannot erase it
bReady := FALSE;                          // 预置未就绪 / preset not ready
nErrCode := 0;                            // 预置无错误码 / preset no error code
bError := FALSE;                          // 预置无故障标志 / preset no fault flag
bValid := TRUE;                           // 预置输出可用 / preset outputs valid
IF _eState = E_DL_BrakeRelState.eFault THEN
    nErrCode := _uErrLatch;               // 重发布锁存故障码，HMI 不会看到码位闪断 / republish the latched fault code
    bError := TRUE;                       // 故障态恒置故障标志 / fault flag stays raised in the fault state
    bValid := FALSE;                      // 故障态输出不可信 / outputs not valid in the fault state
END_IF

// 段 3｜参数与采样门禁：非法即锁存故障并转 eFault，不进状态机（已在故障态则不覆盖原锁存码）
// segment 3, parameter and sample gate; any violation latches a fault and jumps to eFault, an existing latch is not overwritten
_bGateOk := (fReleaseTh > DL_BRI_ZERO) AND (tTorqueQual > DL_BRI_T_ZERO)
        AND (tReleaseTimeout > DL_BRI_T_ZERO) AND (tCloseWait > DL_BRI_T_ZERO);
IF (fTorque <> fTorque) OR ((fTorque - fTorque) <> (fTorque - fTorque)) THEN
    _bGateOk := FALSE;                    // 力矩采样 NaN 或 ±Inf，非有限判定 / torque sample NaN or infinite
END_IF
IF (NOT _bGateOk) AND (_eState <> E_DL_BrakeRelState.eFault) THEN
    IF (fTorque <> fTorque) OR ((fTorque - fTorque) <> (fTorque - fTorque)) THEN
        _uErrLatch := 16#0005_1D04;       // 锁存采样非有限码 / latch the non-finite sample code
        nErrCode := 16#0005_1D04;         // 故障级码赋值 3 行内置 bError / fault-class assignment with bError inline
        bError := TRUE;
        bValid := FALSE;
    ELSE
        _uErrLatch := 16#0005_1D05;       // 锁存参数非法码 / latch the illegal parameter code
        nErrCode := 16#0005_1D05;         // 故障级码赋值 3 行内置 bError / fault-class assignment with bError inline
        bError := TRUE;
        bValid := FALSE;
    END_IF
    _eState := E_DL_BrakeRelState.eFault; // 直接转故障，本拍 CASE 按 eFault 分派 / jump to fault, CASE dispatches on eFault this scan
END_IF

// 段 4｜主状态机：CASE + ELSE 兜底；每个相注明 拍 N 进入 / 本拍行为 / 拍 N+1 转出
// segment 4, main state machine, CASE with ELSE fallback; each phase notes entry, per-scan behaviour and exits
CASE _eState OF
E_DL_BrakeRelState.eIdle:
    // 拍 N 进入：复位后或回闸完成；本拍行为：全失电等待；拍 N+1 转出：使能建立 → eTorqueQual
    // entered after reset or re-close; idle with outputs off; exits to eTorqueQual when the enable appears
    IF bServoEnabled THEN
        _bLostInReady := FALSE;           // 新序默认按中途丢失口径 / new sequence defaults to the mid-sequence class
        _eState := E_DL_BrakeRelState.eTorqueQual; // 进力矩确认相，下一拍计时启动 / enter torque qualification, timing starts next scan
    END_IF

E_DL_BrakeRelState.eTorqueQual:
    // 拍 N 进入：使能建立；本拍行为：力矩低于阈值则 fbTorqueQual 计时；拍 N+1 转出三路：
    // 计时到 → eReleasing；使能丢失 → eClosing（1D03）；门禁非法 → eFault（段 3 已转）
    // entered on enable; timer runs while torque is under threshold; exits to eReleasing on Q,
    // to eClosing on enable loss (1D03), or to eFault via the segment-3 gate
    IF NOT bServoEnabled THEN
        _bLostInReady := FALSE;           // 中途丢失，eClosing 发布 1D03 / lost mid-sequence, eClosing publishes 1D03
        _eState := E_DL_BrakeRelState.eClosing; // 回闸相，输出映射本拍即撤命令 / re-close phase, command drops this scan
    ELSIF fbTorqueQual.Q THEN
        _eState := E_DL_BrakeRelState.eReleasing; // 力矩确认通过，发释放命令 / torque qualified, assert the release command
    END_IF

E_DL_BrakeRelState.eReleasing:
    // 拍 N 进入：力矩确认通过；本拍行为：命令保持、等反馈；拍 N+1 转出三路：
    // 反馈到位 → eReady；超时 → eFault（1D01）；使能丢失 → eClosing（1D03）
    // entered after torque qualification; command held awaiting feedback; exits to eReady on feedback,
    // to eFault on timeout (1D01), or to eClosing on enable loss (1D03)
    IF NOT bServoEnabled THEN
        _bLostInReady := FALSE;           // 中途丢失，eClosing 发布 1D03 / lost mid-sequence, eClosing publishes 1D03
        _eState := E_DL_BrakeRelState.eClosing; // 立即回闸，先于一切确认 / re-close at once, before any acknowledgement
    ELSIF bBrakeReleased THEN
        _eState := E_DL_BrakeRelState.eReady;   // 反馈确认，互锁放行 / feedback confirmed, interlock passes
    ELSIF fbReleaseTo.Q THEN
        _uErrLatch := 16#0005_1D01;       // 锁存反馈超时码 / latch the feedback timeout code
        nErrCode := 16#0005_1D01;         // 故障级码赋值 3 行内置 bError / fault-class assignment with bError inline
        bError := TRUE;
        bValid := FALSE;
        _eState := E_DL_BrakeRelState.eFault;   // 撤输出回退，弹簧闸抱死为安全侧 / roll back, spring brake engagement is the safe side
    END_IF

E_DL_BrakeRelState.eReady:
    // 拍 N 进入：释放反馈确认；本拍行为：命令保持、就绪置位（输出映射段）；拍 N+1 转出两路：
    // 使能丢失 → eClosing（1D02，立即重新上闸）；反馈意外跌落 → eFault（1D06）
    // entered on release feedback; command held and ready asserted; exits to eClosing on enable loss (1D02),
    // or to eFault when the feedback drops unexpectedly (1D06)
    IF NOT bBrakeReleased THEN
        _uErrLatch := 16#0005_1D06;       // 锁存反馈意外跌落码 / latch the unexpected feedback drop code
        nErrCode := 16#0005_1D06;         // 故障级码赋值 3 行内置 bError / fault-class assignment with bError inline
        bError := TRUE;
        bValid := FALSE;
        _eState := E_DL_BrakeRelState.eFault;   // 非受控闭合必须停机检查 / uncontrolled engagement demands a stop
    ELSIF NOT bServoEnabled THEN
        _bLostInReady := TRUE;            // 就绪态丢失，eClosing 发布 1D02 / lost in ready, eClosing publishes 1D02
        _eState := E_DL_BrakeRelState.eClosing; // 立即重新上闸 / re-apply the brake at once
    END_IF

E_DL_BrakeRelState.eClosing:
    // 拍 N 进入：任一相使能丢失；本拍行为：命令已撤、按丢失口径发布信息码、等闭合确认；
    // 拍 N+1 转出：反馈闭合或 tCloseWait 兜底到 → eIdle
    // entered on enable loss from any phase; command off, info code published per class, awaiting closure;
    // exits to eIdle on closed feedback or the tCloseWait fallback
    IF _bLostInReady THEN
        nErrCode := 16#0005_1D02;         // 信息级：就绪态丢使能已回闸，不置 bError / info class, no fault flag
    ELSE
        nErrCode := 16#0005_1D03;         // 信息级：时序中途丢使能已回闸 / info class for the mid-sequence loss
    END_IF
    IF (NOT bBrakeReleased) OR fbCloseWait.Q THEN
        _eState := E_DL_BrakeRelState.eIdle;    // 闸已确认闭合（或时间兜底）回待机 / brake confirmed closed, back to idle
    END_IF

E_DL_BrakeRelState.eFault:
    // 拍 N 进入：任一故障级路径；本拍行为：命令保持撤销、锁存码回放；拍 N+1 转出：
    // bReset 上升沿且无使能 → eIdle（带使能复位禁止，防止立即重新放闸）
    // entered from any fault path; command stays off and the latch replays; exits to eIdle only on
    // a reset edge with no servo enable, so the brake cannot release again immediately
    IF rtReset.Q AND (NOT bServoEnabled) THEN
        _uErrLatch := 0;                  // 清锁存码 / clear the latched code
        _eState := E_DL_BrakeRelState.eIdle;    // 回待机，等下一次使能建立 / back to idle for the next enable
    END_IF

ELSE
    // 非法状态拦截：任何未定义枚举值一律锁存兜底码并转故障（R6）
    // illegal-state interception, any undefined enum value latches the fallback code and goes to fault
    _uErrLatch := 16#0005_1D07;           // 锁存兜底码 / latch the fallback code
    nErrCode := 16#0005_1D07;             // 故障级码赋值 3 行内置 bError / fault-class assignment with bError inline
    bError := TRUE;
    bValid := FALSE;
    _eState := E_DL_BrakeRelState.eFault;
END_CASE

// 段 5｜输出映射：命令只在 eReleasing/eReady 保持，其余相（含故障）一律撤销
// segment 5, output map; the command is held only in eReleasing/eReady and dropped everywhere else including fault
bBrakeReleaseCmd := (_eState = E_DL_BrakeRelState.eReleasing)
                OR (_eState = E_DL_BrakeRelState.eReady); // 释放命令按相映射 / release command mapped by phase
bReady := (_eState = E_DL_BrakeRelState.eReady);          // 就绪仅在确认相 / ready only in the confirmed phase
eState := _eState;                                        // 状态镜像输出 / state mirror output

END_FUNCTION_BLOCK

(* ---- FB_DL_BrakeWearAccum.st ---- *)
(*==============================================================================
 * 组件名称 (Component)  : FB_DL_BrakeWearAccum
 * 所属子库 (Sublibrary) : DL_Motion
 * 当前版本 (Version)    : 1.0.0
 * 兼容性 (Platform)     : CODESYS 3.5+ / TwinCAT 3 / 汇川 InoProShop / 施耐德 Machine Expert
 *                         仅依赖 Standard.library（R_TRIG），零厂商私有库，
 *                         零轴状态枚举引用（R277）
 * 功能描述 (Function)   : 抱闸磨损里程累计。两种磨损源并行累计：① 制动投入
 *                         时长积分（bBrakeOn 电平 × fWearRatePctPerS）；
 *                         ② 投入次数加权（bBrakeOn 上升沿 × fWearPctPerEngage）。
 *                         磨损百分比累计值对 fWearLimitPct 归一输出 fWearPct，
 *                         达预警阈 fWarnPct → bWearWarn 锁存，达限值 →
 *                         bWearAlarm 锁存（维护动作判据）。与 AxisBrakeTest
 *                         分工：本件被动累计，不执行周期试验。
 * 来源标签 (Origin)     : 自研线（IEC 61131-3 标准语义的道莅防御性实现，clean-room）
 * 分工声明 (Pairing)    : BrakeWearAccum（磨损累计，本件）↔ AxisBrakeTest（周期
 *                         试验，既有件）：本件只做投入时长/次数的磨损加权累计
 *                         与阈值告警，不主动试验抱闸、不判抱闸性能（R298 属主
 *                         边界）。
 * 边界语义 (Boundary)   : ① 时长积分用 tScan 引脚步长（组态闸 > 0），上限饱和
 *                         防精度坍缩；
 *                         ② 沿计数回绕防护（DINT 饱和）；
 *                         ③ 预警/告警锁存独立（归因唯一，R190），复位沿一并清；
 *                         ④ 组态闸：磨损率/限值/扫描周期域检查 → 故障锁存；
 *                         ⑤ 监视型无主状态机（R23 公约）。
 * 输出语义 (Fallback)   : 【R191】bEnable = FALSE → 累计冻结（磨损台账是资产，
 *                         不清零），告警锁存保持；eFault 相 → 冻结 + bError。
 * 码位     (Codes)      : 按 R297 范式零 16# 码位硬编码；错误出口 BOOL(bError)+
 *                         eCause 枚举，码位待主控收口统一派号。
 * 红线自检 (Redline)    : 7 项红线已自检：R1 零全局 ✓｜R2 零物理地址 ✓｜R3 纯 IEC ✓
 *                         R4 饱和防回绕/组态闸 ✓｜R5 双语同行注释 ✓
 *                         R6 N/A（监视型无状态机）✓｜R7 R_TRIG 段 0 无条件刷新 ✓
 * 验收向量 (Acceptance) : V1 fWearRatePctPerS=0.001，投入 100s → fWearPct=0.1；
 *                         V2 每次投入加权 0.01，投入 50 次 → 累计 +0.5；
 *                         V3 fWarnPct=80，fWearLimitPct=100 → 80 时 bWearWarn，
 *                         100 时 bWearAlarm（独立锁存）；
 *                         V4 复位沿全清（台账归零语义，上电回夹防线）。
 * 修订历史 (Revision)   : 2026-11-20  v1.0.0  R49 首版（批 4 · 序号 20）
 *==============================================================================*)
TYPE E_DL_BwaCause :
(
    eNone       := 0,                        (* 无故障成因 / No cause *)
    eCfgIllegal := 1                        (* 组态非法：磨损率/限值/周期越域 / Illegal config *)
);
END_TYPE

FUNCTION_BLOCK FB_DL_BrakeWearAccum
VAR_INPUT
    bBrakeOn        : BOOL := FALSE;         (* 制动投入电平（抱闸闭合反馈直连）[-] / Brake-on level *)
    fWearRatePctPerS: LREAL := 0.001;        (* 投入时长磨损率，域 > 0.0 [pct/s] / Wear rate per second *)
    fWearPctPerEngage: LREAL := 0.01;        (* 单次投入磨损加权，域 >= 0.0 [pct/次] / Wear per engagement *)
    fWarnPct        : LREAL := 80.0;         (* 预警阈值，域 0..限值 [pct] / Warning threshold *)
    fWearLimitPct   : LREAL := 100.0;        (* 磨损限值（寿命终点），域 > 预警阈 [pct] / Wear limit *)
    tScan           : TIME := T#10MS;        (* 扫描周期（时长积分步长），域 > T#0S [ms] / Scan cycle step *)
    bEnable         : BOOL := TRUE;          (* 累计使能，FALSE 冻结台账 [-] / Enable *)
    bReset          : BOOL := FALSE;         (* 复位命令，上升沿全清台账与告警锁存 [-] / Reset command *)
END_VAR
VAR_OUTPUT
    fWearPct   : LREAL;                      (* 磨损累计百分比（对限值归一前）[pct] / Accumulated wear percent *)
    fOnTimeS   : LREAL;                      (* 制动投入总时长（台账）[s] / Total brake-on time *)
    nEngageCnt : DINT;                       (* 制动投入总次数（台账）[次] / Total engagement count *)
    bWearWarn  : BOOL;                       (* 达预警阈锁存位（复位沿清）[-] / Wear warning latch *)
    bWearAlarm : BOOL;                       (* 达限值锁存位（复位沿清，独立归因 R190）[-] / Wear alarm latch *)
    eCause     : E_DL_BwaCause;              (* 成因出口（R190 归因唯一） / Cause outlet *)
    bError     : BOOL;                       (* 组态故障锁存标志 [-] / Config fault flag *)
END_VAR
VAR
    rtOn     : R_TRIG;                       (* 投入上升沿实例，段 0 无条件调用 / Engagement edge instance *)
    rtReset  : R_TRIG;                       (* 复位沿实例，段 0 无条件调用 / Reset edge instance *)
    _fWear   : LREAL;                        (* 磨损累计器（锁存量）[pct] / Wear accumulator *)
    _fOnT    : LREAL;                        (* 投入时长累计器（锁存量）[s] / On-time accumulator *)
    _fScanS  : LREAL;                        (* 扫描周期秒值缓存 [s] / Scan seconds cache *)
    _nEng    : DINT;                         (* 投入次数累计器（锁存量）[次] / Engagement counter *)
    _bFault  : BOOL;                         (* 组态故障锁存位 / Config fault latch bit *)
END_VAR
VAR CONSTANT
    DL_BWA_EPS   : LREAL := 1.0E-9;          (* 判零容差 [pct] / Zero epsilon *)
    DL_BWA_SUMMAX: LREAL := 1.0E12;          (* 时长/累计饱和上限（防精度坍缩）[s|pct] / Accumulator saturation *)
    DL_BWA_ENGMAX: DINT  := 1073741824;      (* 次数饱和上限 2^30（防回绕）[次] / Engagement saturation *)
END_VAR

(* —— 段 0：沿实例无条件刷新（R228A） —— *)
rtOn(CLK := bBrakeOn);                       (* 投入沿每拍必调 / On edge every scan *)
rtReset(CLK := bReset);                      (* 复位沿每拍必调 / Reset edge every scan *)

(* —— 段 1：组态闸故障锁存（全引脚覆盖含 NaN 自反，R151/R28；锁存至复位沿，R189） —— *)
IF ((fWearRatePctPerS <= DL_BWA_EPS) OR (fWearPctPerEngage < 0.0)
    OR (fWarnPct < 0.0) OR (fWarnPct > fWearLimitPct) OR (fWearLimitPct <= DL_BWA_EPS)
    OR (tScan <= T#0S)
    OR (fWearRatePctPerS <> fWearRatePctPerS) OR (fWearLimitPct <> fWearLimitPct)) AND NOT _bFault THEN
    _bFault := TRUE;                         (* 组态非法锁存（R45 配对） / Latch config fault *)
    eCause := E_DL_BwaCause.eCfgIllegal;     (* 成因：组态非法 / Cause: illegal config *)
END_IF
_fScanS := TIME_TO_LREAL(tScan) / 1000.0;    (* 毫秒口径换算秒（整毫秒无损）[s] / Convert ms to seconds *)

(* —— 段 2：复位沿处理（作用域：清故障 + 清磨损/时长/次数累计器 + 清双告警锁存，R283 逐项声明） —— *)
IF rtReset.Q THEN
    _bFault := FALSE;                        (* 清故障锁存 / Clear fault *)
    eCause := E_DL_BwaCause.eNone;           (* 清成因 / Clear cause *)
    _fWear := 0.0;                           (* 清磨损累计 / Clear wear *)
    _fOnT := 0.0;                            (* 清时长累计 / Clear on-time *)
    _nEng := 0;                              (* 清次数累计 / Clear count *)
    bWearWarn := FALSE;                      (* 清预警锁存 / Clear warning *)
    bWearAlarm := FALSE;                     (* 清告警锁存 / Clear alarm *)
    fWearPct := 0.0;                         (* 清磨损出口 / Clear wear outlet *)
    fOnTimeS := 0.0;                         (* 清时长出口 / Clear time outlet *)
    nEngageCnt := 0;                         (* 清次数出口 / Clear count outlet *)
END_IF

(* —— 段 3：磨损双源累计（监视型纯派生，无 CASE 相） —— *)
IF bEnable AND NOT _bFault THEN
    IF bBrakeOn THEN
        IF _fOnT < DL_BWA_SUMMAX THEN        (* 时长饱和防护（防精度坍缩） / On-time saturation *)
            _fOnT := _fOnT + _fScanS;        (* 投入时长积分 / On-time integrate *)
        END_IF
        IF _fWear < DL_BWA_SUMMAX THEN       (* 磨损饱和防护 / Wear saturation *)
            _fWear := _fWear + fWearRatePctPerS * _fScanS;   (* 时长磨损加权累计（除法无涉，乘法直算） / Time-based wear accumulate *)
        END_IF
    END_IF
    IF rtOn.Q THEN                           (* 投入沿：次数加权磨损（沿消费已武装，R305） / Engagement edge *)
        IF _nEng < DL_BWA_ENGMAX THEN
            _nEng := _nEng + 1;              (* 次数递增（回绕防护） / Count advance *)
        END_IF
        _fWear := _fWear + fWearPctPerEngage;   (* 次数磨损加权累计 / Engagement wear accumulate *)
    END_IF
    IF _fWear > DL_BWA_SUMMAX THEN
        _fWear := DL_BWA_SUMMAX;             (* 磨损累计兜底饱和 / Wear cap *)
    END_IF
    IF _fWear >= fWearLimitPct THEN
        bWearAlarm := TRUE;                  (* 达限告警锁存至复位沿（独立归因，R190） / Alarm latch *)
    END_IF
    IF _fWear >= fWarnPct THEN
        bWearWarn := TRUE;                   (* 达预警锁存至复位沿（独立归因，R190） / Warning latch *)
    END_IF
END_IF

(* —— 段 4：出口映射（R191 名实同源） —— *)
fWearPct := _fWear;                          (* 磨损出口镜像 / Wear mirror *)
fOnTimeS := _fOnT;                           (* 时长出口镜像 / Time mirror *)
nEngageCnt := _nEng;                         (* 次数出口镜像 / Count mirror *)
bError := _bFault;                           (* 组态故障镜像 / Config fault mirror *)
END_FUNCTION_BLOCK

(* ---- FB_DL_CamFollowerLagMonitor.st ---- *)
(*==============================================================================
 * 组件名称 (Component)  : FB_DL_CamFollowerLagMonitor
 * 所属子库 (Sublibrary) : DL_Motion
 * 当前版本 (Version)    : 1.0.0
 * 兼容性   (Platform)   : CODESYS 3.5+ / TwinCAT 3 / 汇川 InoProShop / 施耐德 Machine Expert
 *                         仅依赖 Standard.library（TON / R_TRIG / ABS），零厂商私有库
 * 功能描述 (Function)   : 凸轮从动轴跟随滞后监控（主从位置差滑动窗统计）。
 *                         每拍采样滞后量 x = fPosMaster − fPosSlave，压入长度 nWindowSize 的
 *                         环形缓冲；每拍在窗内算两个统计量：窗口均值 fLagMean（系统性滞后/超前）
 *                         与窗口内最大绝对值 fLagMax（瞬时最坏滞后）。两档判定：
 *                           预警：|fLagMean| > fLagWarn 或 fLagMax > fLagWarn（维护级，当拍量）
 *                           报警：|fLagMean| > fLagAlarm 或 fLagMax > fLagAlarm，且持续
 *                                 tConfirm（故障锁存）
 *                         均值与最大值并列，是因为二者刻画不同失效：均值大 = 从动轴系统性跟不上
 *                         （增益/惯量问题），最大值大而均值小 = 局部卡顿（机械卡点、润滑不良）。
 *                         只看一个会漏掉另一类故障。
 * 接口     (Interface)  : 输入 fPosMaster 主轴位置、fPosSlave 从动轴位置、nWindowSize 窗长
 *                         （2..64）、fLagWarn / fLagAlarm 阈值、tConfirm 报警确认时间、bReset 复位；
 *                         输出 fLagMean 窗均值、fLagMax 窗最大绝对值、fLagNow 当拍滞后、nFilled
 *                         窗已填数、bWarn 预警、bAlarm 报警锁存、eState / eCause / bError。
 * 边界     (Boundary)   : ① **属主边界（写死）：本件只监控滞后，不输出任何补偿/前馈量，不修改
 *                         凸轮表，不改从动轴指令**。凸轮相位补偿与从动轴前馈属 `FB_DL_ElectronicCam`
 *                         一族；本件的结论位仅供上层做降速/报警/维护决策。
 *                         ② 组态闸：nWindowSize < 2 或 > 64（越 ARRAY 边界）、fLagWarn <= 0.0、
 *                         fLagAlarm <= fLagWarn、tConfirm <= T#0S、位置或阈值 NaN → 故障锁存，
 *                         统计量出口置 0（不宣称）。
 *                         ③ 环形缓冲的窗口统计每拍 O(nWindowSize) 遍历（最大 64 次比较）：
 *                         1 ms 任务下为 64 次浮点比较，可接受；若任务更快请调小 nWindowSize。
 *                         该代价写死在此，不由调用方猜测。
 *                         ④ TON 一枚 + R_TRIG 一枚段 0 无条件周期刷新。
 *                         ⑤ 故障相迁出唯一路径 = bReset 上升沿（R228B）。
 *                         ⑥ 零全局耦合（无 GVL / 无 VAR_EXTERNAL / 无物理地址）。
 * 分工声明 (Scope)      : 与 `FB_DL_AxisFollowingErrorMonitor`（单轴跟随误差）分工——那件比
 *                         "指令位置 vs 实际位置"（同一根轴的指令执行质量），本件比"主轴 vs 从动轴"
 *                         （两根轴之间的相位关系）。电子凸轮下二者都需监控，但归因不同。
 * 来源标签 (Source Tag) : T1-6 ◐（开源参考：凸轮跟随滞后滑动窗统计参数域，零代码行复制）
 * 解除式   (Release)    : bReset 上升沿 ∧ 组态合法 ∧ 当拍 |fLagMean| <= fLagWarn ∧
 *                         当拍 fLagMax <= fLagWarn（R240 全当拍量）。自证可满足：主从追平即满足。
 * 码表     (Codes)      : 本件不占用任何全局数字码位。出口为 REAL 统计量 + BOOL（bWarn / bAlarm /
 *                         bError）+ ENUM（eState / eCause）；数字码位待主控收口阶段统一派号。
 * 红线自检 (Redline)    : R1 ✓ 零 GVL/VAR_EXTERNAL ｜ R2 ✓ 零 %I/%Q/%M ｜ R3 ✓ 纯 IEC 61131-3
 *                         R4 ✓ 数组边界闸 + 阈值几何闸 + 浮点容差 ｜ R5 ✓ 声明逐行同行双语注释
 *                         R6 ✓ ENUM+CASE 含 ELSE ｜ R7 ✓ TON/R_TRIG 段 0 无条件刷新
 * 修订历史 (Revision)   : 2026-11-19  v1.0.0  R46 首版（批次 3 · 序号 11）
 *==============================================================================*)

TYPE E_DL_CflState :
(
    eIdle  := 0,    // 窗未填满，统计量暂不宣称 / Window not filled, statistics not claimed
    eRun   := 10,   // 窗口统计运行相 / Windowed statistics running
    eFault := 90    // 报警锁存相 / Alarm latched phase
);
END_TYPE

TYPE E_DL_CflCause :
(
    eNone       := 0,   // 无异常 / No anomaly
    eCfgIllegal := 1,   // 组态非法（窗长越界/阈值倒置/非有限） / Illegal configuration
    eMeanLimit  := 2,   // 窗均值越报警线（系统性滞后） / Mean lag over the alarm line
    ePeakLimit  := 3,   // 窗峰值越报警线（局部卡顿） / Peak lag over the alarm line
    ePhaseBad   := 4    // 非法相位兜底 / Illegal phase fallback
);
END_TYPE

FUNCTION_BLOCK FB_DL_CamFollowerLagMonitor
VAR_INPUT
    fPosMaster  : REAL := 0.0;      // 主轴位置 [mm] / Master position [mm]
    fPosSlave   : REAL := 0.0;      // 从动轴位置 [mm] / Follower position [mm]
    nWindowSize : INT := 16;        // 滑动窗长度，域 2..64 / Sliding window length, 2..64
    fLagWarn    : REAL := 0.5;      // 滞后期望线，域 > 0.0 [mm] / Lag warning line, > 0.0 [mm]
    fLagAlarm   : REAL := 2.0;      // 滞后报警线，域 > fLagWarn [mm] / Lag alarm line, > warning [mm]
    tConfirm    : TIME := T#100MS;  // 报警确认时间，域 > T#0S [ms] / Alarm confirm time, > 0 [ms]
    bReset      : BOOL := FALSE;    // 复位，上升沿清报警锁存 [-] / Reset, rising edge clears the alarm latch
END_VAR
VAR_OUTPUT
    fLagNow  : REAL;                // 当拍滞后量（主轴 − 从动轴，带符号） [mm] / Present lag, master minus follower [mm]
    fLagMean : REAL;                // 窗口内滞后均值（带符号） [mm] / Windowed mean lag, signed [mm]
    fLagMax  : REAL;                // 窗口内滞后最大绝对值 [mm] / Windowed maximum absolute lag [mm]
    nFilled  : INT;                 // 窗口已填样本数 [个] / Samples currently in the window
    bWarn    : BOOL;                // 维护级预警（未达报警） [-] / Maintenance warning below alarm
    bAlarm   : BOOL;                // 报警锁存 [-] / Latched alarm
    eState   : E_DL_CflState;       // 状态出口 [-] / State outlet
    eCause   : E_DL_CflCause;       // 成因出口（R190 归因唯一） [-] / Cause outlet
    bError   : BOOL;                // 故障标志（报警或组态非法） [-] / Error flag
END_VAR
VAR
    _eState  : E_DL_CflState := E_DL_CflState.eIdle;    // 内部相位（CASE 唯一写入目标） / Internal phase
    _eCause  : E_DL_CflCause := E_DL_CflCause.eNone;    // 成因锁存量 / Latched cause
    tonAlarm : TON;                 // 报警确认计时，段 0 无条件调用 / Alarm confirm timer
    rtReset  : R_TRIG;              // 复位沿实例，段 0 无条件调用 / Reset edge instance
    afRing   : ARRAY[0..63] OF REAL;    // 滞后环形缓冲（64 槽定长，按 nWindowSize 截取） [mm] / Lag ring buffer, fixed 64 slots
    nIdx     : INT;                 // 环形写指针（锁存量） / Ring write index, latched
    nFill    : INT;                 // 已填槽数（锁存量） / Slots filled, latched
    fSum     : REAL;                // 窗内滞后和（锁存量，增量维护） [mm] / Windowed sum, incrementally maintained
    _bFault  : BOOL;                // 报警锁存位（锁存量） / Latched alarm bit
    _bCfgBad : BOOL;                // 组态非法当拍量 [-] / Illegal configuration this scan
    _bNonFin : BOOL;                // 输入非有限当拍量 [-] / Non-finite input this scan
    _fLag    : REAL;                // 当拍滞后中间量 [mm] / Present lag intermediate [mm]
    _fMax    : REAL;                // 窗内最大绝对值中间量 [mm] / Windowed maximum intermediate [mm]
    _fMean   : REAL;                // 窗均值中间量 [mm] / Windowed mean intermediate [mm]
    _i       : INT;                 // 遍历索引 / Loop index
    _bMeanOver : BOOL;              // 均值越报警线当拍量 [-] / Mean over the alarm line
    _bPeakOver : BOOL;              // 峰值越报警线当拍量 [-] / Peak over the alarm line
END_VAR
VAR CONSTANT
    DL_CFL_EPS   : REAL := 1.0E-6;  // 浮点判零容差 [无量纲] / Float epsilon
    DL_CFL_MAXN  : INT := 64;       // 环形缓冲容量（与 afRing 上界一致） [个] / Ring capacity matching afRing bounds
    DL_CFL_MINN  : INT := 2;        // 窗口最小长度（少于 2 无离散意义） [个] / Minimum window length
END_VAR

(* —— 段 0：判据派生 + 两实例无条件周期刷新 —— *)
_bNonFin := (fPosMaster <> fPosMaster) OR (fPosSlave <> fPosSlave)      // NaN 自反判（判等禁令唯一例外） / NaN self-reflexive tests
         OR (fLagWarn <> fLagWarn) OR (fLagAlarm <> fLagAlarm);         // 阈值 NaN 判 / Threshold NaN tests
_bCfgBad := (nWindowSize < DL_CFL_MINN) OR (nWindowSize > DL_CFL_MAXN)  // 窗长越 ARRAY 边界闸 / Window length against array bounds
         OR (fLagWarn <= 0.0) OR (fLagAlarm <= fLagWarn)                // 阈值几何闸 / Threshold geometry gate
         OR (tConfirm <= T#0S) OR _bNonFin;                             // 时间闸 + 非有限 / Time gate and non-finite
_fLag := fPosMaster - fPosSlave;                                        // 当拍滞后（主轴 − 从动轴） / Present lag
rtReset(CLK := bReset);                                                 // 复位沿，每拍必调（R228A） / Reset edge, every scan

(* —— 段 1：单拍量预清零（锁存量 nIdx/nFill/fSum/_bFault/_eCause 不入清单，R107） —— *)
fLagNow := 0.0;         // 当拍滞后出口预清 / Present lag preset
fLagMean := 0.0;        // 均值出口预清 / Mean preset
fLagMax := 0.0;         // 峰值出口预清 / Peak preset
nFilled := 0;           // 填充数出口预清 / Filled preset
bWarn   := FALSE;       // 预警位预清 / Warning preset
bAlarm  := FALSE;       // 报警出口预清 / Alarm preset
bError  := FALSE;       // 故障标志预清（R45 配对） / Error flag preset

(* —— 段 2：复位沿 + 组态闸 —— *)
IF rtReset.Q THEN
    _bFault := FALSE;                                       // 清报警锁存 / Clear alarm latch
    _eCause := E_DL_CflCause.eNone;                         // 清成因 / Clear cause
    nIdx    := 0;                                           // 环形写指针归零 / Ring index cleared
    nFill   := 0;                                           // 填充数归零 / Fill count cleared
    fSum    := 0.0;                                         // 窗口和归零 / Window sum cleared
    IF _eState = E_DL_CflState.eFault THEN
        _eState := E_DL_CflState.eIdle;                     // 故障相迁出（R228B） / Leave fault phase
    END_IF
END_IF
IF _bCfgBad THEN
    _bFault := TRUE;                                        // 组态非法锁存 / Latch illegal configuration
    _eCause := E_DL_CflCause.eCfgIllegal;                   // 归因：组态非法 / Cause: illegal configuration
END_IF

(* —— 段 3：环形缓冲写入（先减被覆盖的旧值，再加新值，保持 fSum 与窗内一致） —— *)
IF NOT _bCfgBad THEN
    IF nFill >= nWindowSize THEN
        fSum := fSum - afRing[nIdx];                        // 覆盖前减掉旧样本 / Subtract the evicted sample
    ELSE
        nFill := nFill + 1;                                 // 窗口未满则填充数增 / Grow the fill count
    END_IF
    afRing[nIdx] := _fLag;                                  // 写入当拍样本 / Store the present sample
    fSum := fSum + _fLag;                                   // 加上新样本 / Add the new sample
    nIdx := nIdx + 1;                                       // 指针前进 / Advance the pointer
    IF nIdx >= nWindowSize THEN
        nIdx := 0;                                          // 到窗长回卷 / Wrap at the window length
    END_IF
    IF nIdx > DL_CFL_MAXN - 1 THEN
        nIdx := 0;                                          // 双保险：绝不让指针越 ARRAY 上界 / Second guard, never index past the array
    END_IF
    IF nFill > nWindowSize THEN
        nFill := nWindowSize;                               // 钳位（窗长改小时自愈） / Clamp when the window shrinks
    END_IF
END_IF

(* —— 段 4：窗口统计（均值与最大绝对值，均在窗内 nFill 个样本上算） —— *)
IF (NOT _bCfgBad) AND (nFill > 0) THEN
    _fMean := fSum / INT_TO_REAL(nFill);                    // 均值，分母已判正（nFill > 0） / Mean, denominator guarded
    _fMax  := 0.0;                                          // 最大值初值 / Peak initial value
    FOR _i := 0 TO nFill - 1 DO
        IF ABS(afRing[_i]) > _fMax THEN
            _fMax := ABS(afRing[_i]);                       // 逐个比较取最大绝对值 / Track the maximum absolute value
        END_IF
    END_FOR
    fLagNow  := _fLag;                                      // 当拍滞后出口 / Present lag outlet
    fLagMean := _fMean;                                     // 均值出口 / Mean outlet
    fLagMax  := _fMax;                                      // 峰值出口 / Peak outlet
    nFilled  := nFill;                                      // 填充数出口 / Filled outlet
END_IF

(* —— 段 5：分档判据（双口径取或；先算判据再喂 TON，保证 IN 由当拍表达式派生） —— *)
_bMeanOver := ((NOT _bCfgBad) AND (nFill > 0)) AND (ABS(fLagMean) > fLagAlarm);     // 均值越报警线 / Mean over the alarm line
_bPeakOver := ((NOT _bCfgBad) AND (nFill > 0)) AND (fLagMax > fLagAlarm);           // 峰值越报警线 / Peak over the alarm line
tonAlarm(IN := _bMeanOver OR _bPeakOver, PT := tConfirm);                           // 报警确认窗 / Alarm confirm window

(* —— 段 6：报警锁存与归因（均值优先于峰值：系统性滞后比局部卡顿更需要先看） —— *)
IF (NOT _bFault) AND (NOT _bCfgBad) AND tonAlarm.Q THEN
    _bFault := TRUE;                                        // 锁存 / Latch
    IF _bMeanOver THEN
        _eCause := E_DL_CflCause.eMeanLimit;                // 归因：均值越限 / Cause: mean over limit
    ELSE
        _eCause := E_DL_CflCause.ePeakLimit;                // 归因：峰值越限 / Cause: peak over limit
    END_IF
END_IF

(* —— 段 7：预警（维护级；报警相不再宣称预警） —— *)
IF (NOT _bFault) AND (NOT _bCfgBad) AND (nFill > 0)
   AND ((ABS(fLagMean) > fLagWarn) OR (fLagMax > fLagWarn)) THEN
    bWarn := TRUE;                                          // 维护级预警 / Maintenance warning
END_IF

(* —— 段 8：锁存相位迁移闸 —— *)
IF _bFault AND (_eState <> E_DL_CflState.eFault) THEN
    _eState := E_DL_CflState.eFault;                        // 锁存即入故障相 / Latch enters fault phase
END_IF

(* —— 段 9：相位机（ENUM 全成员显式标签 + ELSE 兜底，R128） —— *)
CASE _eState OF

E_DL_CflState.eIdle:
    IF _bFault THEN                                         // 出口 1：故障锁存 / Fault latched
        _eState := E_DL_CflState.eFault;
    ELSIF (_bCfgBad = FALSE) AND (nFill >= nWindowSize) THEN    // 出口 2：窗已填满，统计可信 / Window filled, statistics trustworthy
        _eState := E_DL_CflState.eRun;
    END_IF

E_DL_CflState.eRun:
    IF _bFault THEN                                         // 出口 1：报警锁存 / Alarm latched
        _eState := E_DL_CflState.eFault;
    ELSIF nFill < nWindowSize THEN                          // 出口 2：窗被清（复位后重填） / Window cleared, refilling
        _eState := E_DL_CflState.eIdle;
    END_IF

E_DL_CflState.eFault:
    ;                                                       // 故障相：仅段 2 复位沿可迁出 / Only the reset edge leaves this phase

ELSE
    _bFault := TRUE;                                        // 非法相位兜底锁存 / Illegal-phase fallback latch
    _eCause := E_DL_CflCause.ePhaseBad;                     // 归因：非法相位 / Cause: illegal phase
    _eState := E_DL_CflState.eFault;                        // 强拉故障相 / Force fault phase

END_CASE

(* —— 段 10：出口单点映射（名实双出口，R191） —— *)
bAlarm := _bFault;                                          // 报警与锁存同源 / Alarm from latch
bError := _bFault OR _bCfgBad;                              // 故障标志 = 锁存或组态非法 / Error = latch or illegal config
IF _bFault THEN
    bWarn := FALSE;                                         // 报警相不宣称「仅预警」 / No warning claim in alarm
END_IF
eState := _eState;                                          // 状态出口 / State outlet
eCause := _eCause;                                          // 成因出口 / Cause outlet

END_FUNCTION_BLOCK
